(* IEC 61131-3 sources: daoli-st-library/DL_Motion (part 11) *)

(* ---- FB_DL_CamOverrideTrim.st ---- *)
(*
  FB_DL_CamOverrideTrim  —  凸轮运行中动态修调（幅值/相位偏置实时叠加）/ In-run cam dynamic override trim
  分类 Category : DL_Motion
  码位 Code     : 16#04_0_A6
  段位说明      : 04_0 段占至 A5，A6 格空穴，本件启用 A6 格
  版本 Version  : 1.0.1
  来源 Source   : t1-6-plcopen — T1-6 行待挖项「凸轮动态修调」落地
  溯源 Origin   : clean-room 实现，未复制任何源码行
  功能 Function : 1) 不重选表、不脱耦：在 FC_DL_CamTableInterp 表插值输出上实时叠加修调；
                  2) 相位偏置 fPhaseTrim：主轴位置先叠加相位偏置再查表（fMasterEff = fMasterPos + fPhaseTrim），
                  周期模式下按 fPeriod 取模回界，非周期模式下越界按表界钳制（bInRange 反映真实界内性）；
                  3) 幅值偏置 fAmpTrim：从轴输出直接叠加（fSlaveTrimmed = fSlavePos + fAmpTrim）；
                  4) bTrimFreeze 电平冻结修调：冻结拍输出纯表值（修调增量记忆保留，解冻即恢复）。
  边界 Boundary : ① 本件只做输出叠加，不写轴命令、不下使能，凸轮耦合本体由上层承载；
                  ② 与 FC_DL_CamTableInterp（表插值原子）与 FB_DL_ElectronicCam（耦合本体）分工明确；
                  ③ 修调量非有限防御：NaN/Inf 保持上次有效修调值（增量语义不突变）；
                  ④ 无 CASE 主状态机（变换型 FB）：无相位迁移，无跨相 TON 复用问题；
                  ⑤ 本件每拍必须调用一次（无定时器/边沿实例，跳拍仅导致输出陈旧，无隐藏状态损坏）。
  依赖 Depends  : I_DL_MotionAxis（注入，不实例化，只读 fPosition）；
                  FC_DL_CamTableInterp（函数调用，aCam 固定上界透传 + uPointCnt 显式点数）；ST_DL_CamPoint（库内既有结构）
  码表 Error codes（本件格 04_0_A6，子码步进 +0x100）:
    16#0004_01A6 信息级：修调量非有限已保持上次有效值（继续输出，不中断）
    16#0004_02A6 信息级：插值件报错码透传（表非法/越界，本件输出钳界表值）
    16#0004_03A6 信息级：冻结使能中（bTrimFreeze = TRUE，输出纯表值）

  修订历史 Revision :
    2026-11-19  v1.0.0  R39 首版（批次 2 · 序号 7）
    2026-11-23  v1.0.1  R75 适配插值件显式点数字段：aCam 改固定上界 ARRAY[1..200]，
                        增输入 uPointCnt 透传（解 VLA 透传 E037）
*)

FUNCTION_BLOCK FB_DL_CamOverrideTrim
VAR_INPUT
    bEnable     : BOOL := FALSE;      // 使能，FALSE 时输出纯表值（修调旁路）/ Enable, FALSE bypasses trim
    bTrimFreeze : BOOL := FALSE;      // 修调冻结，电平有效：冻结拍输出纯表值 [-] / Trim freeze, level active
    fAmpTrim    : REAL := 0.0;        // 幅值偏置 [mm]，直接叠加从轴输出 / Amplitude trim, added to slave output
    fPhaseTrim  : REAL := 0.0;        // 相位偏置 [mm]，叠加主轴位置后查表 / Phase trim, added to master position
    bPeriodic   : BOOL := FALSE;      // 周期模式使能（与插值件同口径透传）/ Periodic mode, passed to interpolator
    fPeriod     : LREAL := 360.0;     // 周期模式主轴周期 [mm]，域 > 0 / Master period for periodic mode
    bReset      : BOOL := FALSE;      // 修调复位，上升沿清修调保持值（重新从 0 起）/ Trim reset, rising edge clears hold
    uPointCnt   : UINT := 100;        // 凸轮表有效点数，域 [2,200]，透传插值件 [点] / Valid table point count, passthrough to interpolator
END_VAR
VAR_OUTPUT
    fSlaveBase    : LREAL;            // 纯表值输出 [mm]（未叠加修调）/ Pure table output without trim
    fSlaveTrimmed : LREAL;            // 修调后从轴输出 [mm] / Trimmed slave output
    bInRange      : BOOL;             // 有效主轴位置在表界内 [-] / Effective master position within table range
    bTrimActive   : BOOL;             // 修调实际生效中（使能且未冻结且偏置非零）/ Trim actually active
    bClampEdge    : BOOL;             // 相位偏置越表界被钳制（非周期模式）/ Phase trim clamped at table edge
    uErrorId      : UDINT;            // 事件码，0 = 无事件（本件码均信息级瞬时）/ Event code, transient info only
END_VAR
VAR_IN_OUT
    iAxis : I_DL_MotionAxis;          // 主轴引用（注入，不实例化，只读位置）/ Master axis reference, position read-only
    aCam  : ARRAY[1..200] OF ST_DL_CamPoint; // 凸轮表透传（固定上界，下标 1..uPointCnt 有效，须按 fMaster 升序）/ Cam table passed through, fixed bound
END_VAR
VAR
    rtReset      : R_TRIG;            // 修调复位沿实例，主体首部无条件刷新 / Trim reset edge instance
    _bInRangeInt : BOOL;              // 插值件表界内标志内部镜像（段 3 每拍接收，直赋出口）[-] / Interp in-range mirror, received every scan in seg 3
    fAmpTrimEff  : REAL := 0.0;       // 生效幅值偏置 [mm]（非有限保持载体）/ Effective amplitude trim with hold
    fPhaseTrimEff: REAL := 0.0;       // 生效相位偏置 [mm]（非有限保持载体）/ Effective phase trim with hold
    fMasterEff   : LREAL;             // 修调后有效主轴位置 [mm] / Effective master position after phase trim
    fSlavePos    : LREAL;             // 插值件从轴输出 [mm] / Interpolator slave output
    eInterpErr   : UDINT;             // 插值件本拍错误码透传 / Interpolator error code passthrough
    bDefend      : BOOL;              // 本拍非有限防御触发标志 / Non-finite defense triggered this cycle
END_VAR
VAR CONSTANT
    DL_COT_INF_CAP : LREAL := 1.0E15;   // 非有限值筛查幅值上限 / Non-finite screening cap
END_VAR

(* —— 段 0：边沿实例无条件周期刷新（R7 红线） —— *)
rtReset(CLK := bReset);                 // 修调复位沿刷新，每拍必调

(* —— 段 1：修调量非有限防御（NaN/Inf 保持上次有效值；复位沿清保持） —— *)
bDefend := FALSE;                       // 防御标志预清零
IF (fAmpTrim <> fAmpTrim) OR (ABS(fAmpTrim) > DL_COT_INF_CAP) OR ((fAmpTrim - fAmpTrim) <> 0.0) THEN
    bDefend := TRUE;                    // 幅值偏置非有限：保持上次有效
ELSE
    fAmpTrimEff := fAmpTrim;            // 有效值入保持载体
END_IF
IF (fPhaseTrim <> fPhaseTrim) OR (ABS(fPhaseTrim) > DL_COT_INF_CAP) OR ((fPhaseTrim - fPhaseTrim) <> 0.0) THEN
    bDefend := TRUE;                    // 相位偏置非有限：保持上次有效
ELSE
    fPhaseTrimEff := fPhaseTrim;        // 有效值入保持载体
END_IF
IF rtReset.Q THEN
    fAmpTrimEff := 0.0;                 // 复位沿：幅值修调归零
    fPhaseTrimEff := 0.0;               // 复位沿：相位修调归零
END_IF

(* —— 段 2：相位偏置叠加（主轴位置先偏置，周期模式取模回界） —— *)
IF bPeriodic AND (fPeriod > 0.0) THEN
    fMasterEff := iAxis.fPosition + fPhaseTrimEff;              // 叠加相位偏置
    fMasterEff := fMasterEff - TRUNC(fMasterEff / fPeriod) * fPeriod;   // 取模回界（分母已闸 > 0）
    IF fMasterEff < 0.0 THEN
        fMasterEff := fMasterEff + fPeriod;                     // 负模回正（保持 [0, fPeriod) 域）
    END_IF
    bClampEdge := FALSE;                                        // 周期模式无表界钳制概念
ELSE
    fMasterEff := iAxis.fPosition + fPhaseTrimEff;              // 非周期：直接叠加（界内性由插值件判）
    bClampEdge := FALSE;                                        // 钳制判定由插值件 bInRange 承载
END_IF

(* —— 段 3：调表插值原子（每拍一次；错误码透传） —— *)
FC_DL_CamTableInterp(fMasterPos := fMasterEff,      // 有效主轴位置（已含相位偏置）
                     bPeriodic := bPeriodic,        // 周期模式透传
                     fPeriod := fPeriod,            // 周期透传
                     uPointCnt := uPointCnt,        // 显式点数透传（R75 口径）/ Explicit point count passthrough
                     aCam := aCam,                  // 凸轮表透传（固定上界数组引用）
                     fSlavePos => fSlavePos,        // 从轴表值输出
                     bInRange => _bInRangeInt,      // 表界内标志输出（内部镜像）/ In-range flag to internal mirror
                     eErr => eInterpErr);           // 插值件错误码输出
fSlaveBase := fSlavePos;                            // 纯表值镜像
bInRange := _bInRangeInt;                           // 表界内标志出口每拍直赋（语义：有效主轴位置在凸轮表界内为 TRUE）/ In-range outlet assigned every scan

(* —— 段 4：幅值修调叠加与使能门控 —— *)
IF bEnable AND (NOT bTrimFreeze) THEN
    fSlaveTrimmed := fSlaveBase + fAmpTrimEff;      // 修调生效：表值 + 幅值偏置
    bTrimActive := (fAmpTrimEff <> 0.0) OR (fPhaseTrimEff <> 0.0);   // 修调非零即生效中
ELSE
    fSlaveTrimmed := fSlaveBase;                    // 旁路/冻结：输出纯表值（修调保持值不丢）
    bTrimActive := FALSE;
END_IF

(* —— 段 5：事件码合成（信息级瞬时，无锁存） —— *)
uErrorId := 16#0000_0000;               // 缺省无事件
IF bDefend THEN
    uErrorId := 16#0004_01A6;           // 信息级：修调量非有限已保持
ELSIF eInterpErr <> 0 THEN
    uErrorId := 16#0004_02A6;           // 信息级：插值件错误码透传
END_IF
IF bTrimFreeze AND bEnable THEN
    uErrorId := 16#0004_03A6;           // 信息级：冻结使能中（覆盖优先级最低，放最后）
END_IF

END_FUNCTION_BLOCK

(* ---- FB_DL_CamPhaseTrim.st ---- *)
(*
    FB_DL_CamPhaseTrim —— 凸轮相位在线修调
    ------------------------------------------------------------------
    分类      : DL_Motion / Cam
    前缀      : FB_DL_
    版本      : 1.0.0
    溯源      : 只借「凸轮相位可在线修调属运动层能力」的公开语义与运动层组织事实；
                限速率渐进、标记沿一次性受理、相位归一的禁 MOD 写法、错误分级与
                码位 100% 自有；本件不自造轴状态、不内联凸轮算法（组合调用上层凸轮件）；
                clean-room 重写，未复制任何闭源厂商源码
    平台      : 纯 IEC 61131-3，CODESYS V3.5+ / TwinCAT 3 / InoProShop 通用
    作者      : 道莅代码库 · PLC编程专家（R19）
    ------------------------------------------------------------------
    功能说明  : 运行中在线修调凸轮相位，输出一个相位偏移量注入凸轮件的相位输入
                （组合而非内联：可依赖低层，但不复制低层）。现场语义是飞剪/横切/贴标的
                切点对位——用色标或标记传感器测到实际相位偏差后一点点修，修的过程必须
                限速率，突变等于给机械一个冲击。
                核心防御：① 相位限幅越域（> 180°）或速率越域即故障级 02E1 并冻结修调——
                   相位限幅 0 会让修调永久卡住、太大等于允许突变；
                ② 一次性标记补偿每标记沿只受理一次，且必须在 bMarkArmed（上一拍已复位）
                   时才受理——否则高频标记会在一拍内累加成大跳变（本件最高危点）；
                ③ 相位归一用条件加减，禁浮点 MOD；
                ④ 指令或补偿量非有限即故障级并保持末次偏移——归 0 会让切点瞬间错位切出废品；
                ⑤ bReset 立即清偏移（唯一允许跳变的路径，检修专用）。
                职责边界：凸轮曲线求值归电子凸轮件，本件只出相位偏移量。
    错误码    : 16#0004_01CF 目标偏移超限已钳位 / 单次标记补偿已生效——信息级，正常防御
                16#0004_01D0 预留禁用（信息级，不得挪用）
                16#0004_02E1 限幅、速率或采样周期参数非法——故障级，修调冻结且偏移保持
                16#0004_02E2 指令或补偿量非有限——故障级，偏移保持末次有效
                16#0004_02E3 状态机落 ELSE 兜底（非法状态）——故障级，回 eIdle 并保持偏移
    码位总账  : 16#0004_01CF 用 / 16#0004_01D0 预留 ｜ 16#0004_02E1 用 / 16#0004_02E2 用 / 16#0004_02E3 用
    状态机    : E_DL_TrimState（eIdle / eRamping / eHold / eFault）四态，CASE 含 ELSE 兜底，
                ELSE 回 eIdle 并置故障级 02E3；失能时目标归 0 并按限速率回零。
    采样约定  : fbTrigReset / fbTrigMark 在本体首部无条件刷新，绝不放入 IF 或 CASE；
                速率步长由 tSampleTime 引脚换算，首拍步长按引脚值直接给出（无历史依赖）。
    修订记录  : 2026-11-16 v1.0.0 首次入库（R19）
*)

(*
    枚举 : E_DL_TrimState —— 相位修调状态（本文件为全库唯一属主）
*)
TYPE E_DL_TrimState :
(
    eIdle    := 0,                            // 空闲：偏移按限速率回零 / idle, the offset ramps back to zero
    eRamping := 1,                            // 趋近：向目标偏移逼近 / ramping towards the target offset
    eHold    := 2,                            // 保持：已到目标，仅受标记补偿影响 / holding at the target
    eFault   := 3                             // 故障：修调冻结，偏移保持 / fault, the trim is frozen and the offset held
);
END_TYPE

FUNCTION_BLOCK FB_DL_CamPhaseTrim
VAR_INPUT
    bEnable         : BOOL;                   // 使能，FALSE 偏移按限速率归 0 / enable, FALSE ramps the offset back to zero
    bReset          : BOOL;                   // 复位，上升沿立即清偏移（检修专用，会跳变）/ reset, rising edge clears the offset at once, maintenance only
    fPhaseOffsetCmd : REAL := 0.0;            // 目标相位偏移 [deg]，范围 -180.0~180.0 / target phase offset [deg], range -180.0~180.0
    fRateMax        : REAL := 30.0;           // 偏移变化率上限 [deg/s]，范围 0.1~3600.0 / maximum offset rate [deg/s], range 0.1~3600.0
    fPhaseLimit     : REAL := 90.0;           // 偏移绝对值上限 [deg]，范围 1.0~180.0 / absolute offset limit [deg], range 1.0~180.0
    bTrimOnMark     : BOOL := FALSE;          // TRUE = 叠加标记沿的一次性补偿 / TRUE adds the one-shot mark correction
    fMarkCorrection : REAL := 0.0;            // 单次标记补偿量 [deg]，范围 -10.0~10.0 / one-shot mark correction [deg], range -10.0~10.0
    bMarkPulse      : BOOL := FALSE;          // 标记传感器脉冲（上升沿有效）/ mark sensor pulse, rising edge valid
    tSampleTime     : TIME := T#10MS;         // 采样周期 [ms]，范围 1~1000 / sample time [ms], range 1~1000
END_VAR
VAR_OUTPUT
    fPhaseOffset    : REAL;                   // 实际输出相位偏移（注入凸轮件）[deg] / actual phase offset injected into the cam block [deg]
    bTrimming       : BOOL;                   // 正在趋近目标 / ramping towards the target
    bLimited        : BOOL;                   // 受速率或幅值限制 / limited by the rate or the magnitude
    uMarkCount      : UDINT;                  // 已受理的标记补偿次数，饱和 [次] / accepted mark corrections, saturating [times]
    eErr            : UDINT;                  // 错误码，0=正常 / error id, 0=ok
    bError          : BOOL;                   // 故障标志，eErr 为故障级时 TRUE / error flag, TRUE on fault-level eErr
END_VAR
VAR
    fbTrigReset     : R_TRIG;                 // 复位上升沿实例，本体首部无条件刷新 / reset edge instance, refreshed unconditionally
    fbTrigMark      : R_TRIG;                 // 标记上升沿实例，本体首部无条件刷新 / mark edge instance, refreshed unconditionally
    eState          : E_DL_TrimState := eIdle; // 状态机当前态 / current state machine state
    fOffset         : REAL;                   // 内部偏移量 [deg] / internal offset [deg]
    fTarget         : REAL;                   // 限幅后的目标偏移 [deg] / clamped target offset [deg]
    fStep           : REAL;                   // 本拍允许的最大变化量 [deg] / maximum allowed change in this cycle [deg]
    fDtSec          : REAL;                   // 采样周期秒值 [s] / sample time in seconds [s]
    fLimitEff       : REAL;                   // 钳位后的相位限幅 [deg] / clamped phase limit [deg]
    fCorrEff        : REAL;                   // 钳位后的单次补偿量 [deg] / clamped one-shot correction [deg]
    bMarkArmed      : BOOL := TRUE;           // 标记受理武装位（上一拍已复位才受理）/ mark acceptance arming bit, armed only after the pulse is released
    bNonFin         : BOOL;                   // 输入非有限判定标志 / non-finite input flag
    bInit           : BOOL := FALSE;          // 首扫标志，初值 FALSE，判据 NOT bInit / first-scan flag, initial FALSE, tested with NOT
    nDtMs           : DINT;                   // 采样周期毫秒整数 [ms] / sample time in integer milliseconds [ms]
END_VAR
VAR CONSTANT
    DL_CPT_LIMIT_MAX : REAL := 180.0;         // 相位限幅上限（半周）[deg] / phase limit upper bound, half a revolution [deg]
    DL_CPT_LIMIT_MIN : REAL := 1.0;           // 相位限幅下限 [deg] / phase limit lower bound [deg]
    DL_CPT_RATE_MAX  : REAL := 3600.0;        // 速率上限 [deg/s] / rate upper bound [deg/s]
    DL_CPT_RATE_MIN  : REAL := 0.1;           // 速率下限 [deg/s] / rate lower bound [deg/s]
    DL_CPT_MARK_MAX  : REAL := 10.0;          // 单次补偿量绝对值上限 [deg] / absolute one-shot correction bound [deg]
    DL_CPT_DT_MAX    : TIME := T#1S;          // 采样周期上限 [ms] / sample time upper bound [ms]
    DL_CPT_DT_MIN    : TIME := T#1MS;         // 采样周期下限 [ms] / sample time lower bound [ms]
    DL_FLOAT_EPS     : REAL := 1.0E-6;        // 浮点判等容差 [无量纲] / float equality tolerance [dimensionless]
    DL_CPT_FULL_TURN : REAL := 360.0;         // 一整周 [deg] / one full revolution [deg]
    DL_CPT_HALF_TURN : REAL := 180.0;         // 半周 [deg] / half a revolution [deg]
    DL_CPT_MS_PER_S  : REAL := 1000.0;        // 毫秒到秒换算因子 [ms/s] / milliseconds per second [ms/s]
    DL_CPT_INF_GUARD : REAL := 1.0E38;        // 非有限幅值判定阈值 [无量纲] / non-finite magnitude guard [dimensionless]
    DL_CPT_CNT_MAX   : UDINT := 16#FFFF_FFFE; // 标记次数饱和值 [次] / mark counter saturation value [times]
    DL_CPT_ZERO      : REAL := 0.0;           // 零值常量，避免裸字面量 [deg] / zero constant, avoids a bare literal [deg]
END_VAR

// 段 1｜边沿实例无条件周期刷新（红线：严禁放入条件分支）/ segment 1, unconditional edge refresh
fbTrigReset(CLK := bReset);
fbTrigMark(CLK := bMarkPulse);

// 段 2｜输出与错误状态预置 / segment 2, preset outputs and status
eErr := 0;                                    // 预置无错误 / preset no error
bError := FALSE;                              // 预置无故障 / preset no fault
bTrimming := FALSE;                           // 预置未趋近 / preset not ramping
bLimited := FALSE;                            // 预置未受限 / preset not limited

// 段 3｜首扫初始化（唯一合法范式：初值 FALSE，判据 NOT bInit）/ segment 3, first-scan initialisation
IF NOT bInit THEN
    fOffset := DL_CPT_ZERO;                   // 首扫偏移归 0，避免未定值上电冲击 / the offset starts at zero, no undefined jump at power up
    uMarkCount := 0;                          // 标记计数清零 / clear the mark counter
    bInit := TRUE;                            // 首扫只做一次 / first scan runs once only
END_IF

// 段 4｜参数闸（限幅、速率、采样周期，任一非法即冻结修调）/ segment 4, parameter gate freezes the trim
IF (fPhaseLimit < DL_CPT_LIMIT_MIN) OR (fPhaseLimit > DL_CPT_LIMIT_MAX)
   OR (fRateMax < DL_CPT_RATE_MIN) OR (fRateMax > DL_CPT_RATE_MAX)
   OR (tSampleTime < DL_CPT_DT_MIN) OR (tSampleTime > DL_CPT_DT_MAX) THEN
    eErr := 16#0004_02E1;                     // 参数非法故障码 / illegal parameter fault id
    bError := TRUE;                           // 置故障标志 / raise the error flag
    eState := eFault;                         // 落故障态，修调冻结 / enter the fault state, the trim is frozen
    fPhaseOffset := fOffset;                  // 偏移保持，绝不归 0 / hold the offset, never reset it to zero
    RETURN;                                   // 故障级提前返回 / early return on fault
END_IF

// 段 5｜输入非有限闸：偏移保持末次有效（归 0 会瞬间错位切出废品）/ segment 5, non-finite gate holds the offset
bNonFin := (fPhaseOffsetCmd <> fPhaseOffsetCmd) OR (fMarkCorrection <> fMarkCorrection)
        OR (fPhaseOffsetCmd > DL_CPT_INF_GUARD) OR (fPhaseOffsetCmd < -DL_CPT_INF_GUARD); // 非有限判定 / non-finite detection
IF bNonFin THEN
    eErr := 16#0004_02E2;                     // 指令非有限故障码 / non-finite command fault id
    bError := TRUE;                           // 置故障标志 / raise the error flag
    eState := eFault;                         // 落故障态 / enter the fault state
    fPhaseOffset := fOffset;                  // 保持末次有效偏移 / hold the last valid offset
    RETURN;                                   // 故障级提前返回 / early return on fault
END_IF

// 段 5｜域钳位（限幅、补偿量各自收敛，钳位本身不置码）/ segment 5, domain clamp
fLimitEff := MIN(MAX(fPhaseLimit, DL_CPT_LIMIT_MIN), DL_CPT_LIMIT_MAX);   // 相位限幅收敛 [deg] / converge the phase limit [deg]
fCorrEff := MIN(MAX(fMarkCorrection, -DL_CPT_MARK_MAX), DL_CPT_MARK_MAX); // 单次补偿收敛到 ±10 deg / converge the one-shot correction
nDtMs := TIME_TO_DINT(tSampleTime);           // 采样周期整数毫秒 [ms] / sample time in integer milliseconds [ms]
fDtSec := DINT_TO_REAL(nDtMs) / DL_CPT_MS_PER_S; // 换算为秒，除子为常量 [s] / convert to seconds, the divisor is a constant [s]
fStep := fRateMax * fDtSec;                   // 本拍允许的最大变化量 [deg] / maximum allowed change in this cycle [deg]

// 段 6｜目标偏移 = 指令限幅 / segment 6, target offset from the clamped command
fTarget := MIN(MAX(fPhaseOffsetCmd, -fLimitEff), fLimitEff); // 目标双侧钳位 [deg] / clamp the target on both sides [deg]
IF ABS(fPhaseOffsetCmd) > fLimitEff THEN
    eErr := 16#0004_01CF;                     // 信息级：目标偏移超限已钳位 / info level, the target was clamped
END_IF

// 段 7｜标记沿一次性补偿（最高危点：每沿只受理一次，且需武装位）/ segment 7, one-shot mark correction
IF NOT bMarkPulse THEN
    bMarkArmed := TRUE;                       // 脉冲释放即重新武装 / re-arm once the pulse is released
END_IF
IF fbTrigMark.Q AND bTrimOnMark AND bMarkArmed THEN
    bMarkArmed := FALSE;                      // 受理后立即解除武装，防同拍累加 / disarm immediately so no accumulation can happen in one cycle
    fTarget := MIN(MAX(fTarget + fCorrEff, -fLimitEff), fLimitEff); // 叠加补偿并限幅 [deg] / add the correction and clamp [deg]
    IF uMarkCount < DL_CPT_CNT_MAX THEN
        uMarkCount := uMarkCount + 1;         // 饱和计数 / saturating count
    END_IF
    eErr := 16#0004_01CF;                     // 信息级：单次标记补偿已生效 / info level, the one-shot correction was applied
END_IF

// 段 8｜复位沿：立即清偏移（唯一允许跳变的路径，检修专用）/ segment 8, reset clears the offset at once
IF fbTrigReset.Q THEN
    fOffset := DL_CPT_ZERO;                   // 检修专用清偏移 / maintenance only, clear the offset
    bLimited := FALSE;                        // 清限幅标志 / clear the limited flag
END_IF

// 段 9｜失能：目标归 0，按限速率回零 / segment 9, disabling ramps the target back to zero
IF NOT bEnable THEN
    fTarget := DL_CPT_ZERO;                   // 目标归 0 / the target returns to zero
END_IF

// 段 10｜状态机（含 ELSE 兜底）/ segment 10, state machine with ELSE fallback
CASE eState OF
    eIdle:
        IF ABS(fTarget - fOffset) > fStep THEN
            eState := eRamping;               // 偏离超过一步即进入趋近态 / a deviation beyond one step enters the ramping state
        ELSE
            eState := eHold;                  // 否则直接保持 / otherwise hold at once
        END_IF

    eRamping:
        IF ABS(fTarget - fOffset) <= fStep THEN
            eState := eHold;                  // 进入一步之内即趋近完成 / inside one step the ramp is finished
        END_IF

    eHold:
        IF ABS(fTarget - fOffset) > fStep THEN
            eState := eRamping;               // 新指令或标记补偿把偏差拉大即重新趋近 / a new command or correction restarts the ramp
        END_IF

    eFault:
        fPhaseOffset := fOffset;              // 故障态偏移保持 / hold the offset in the fault state

ELSE
    eErr := 16#0004_02E3;                     // 故障级：非法状态兜底 / fault level, illegal state fallback
    bError := TRUE;                           // 置故障标志 / raise the error flag
    eState := eIdle;                          // 回空闲态 / fall back to idle
    fPhaseOffset := fOffset;                  // 保持偏移，绝不清零 / hold the offset, never clear it
END_CASE

// 段 11｜限速率推进（每拍最多变化 fStep，禁浮点 MOD 的相位归一）/ segment 11, rate limited advance
IF eState <> eFault THEN
    IF fOffset > (fTarget + fStep) THEN
        fOffset := fOffset - fStep;           // 正向逼近 / approach from above
        bLimited := TRUE;                     // 标记速率受限 / flag the rate limit
        bTrimming := TRUE;                    // 正在趋近 / ramping
    ELSIF fOffset < (fTarget - fStep) THEN
        fOffset := fOffset + fStep;           // 负向逼近 / approach from below
        bLimited := TRUE;                     // 标记速率受限 / flag the rate limit
        bTrimming := TRUE;                    // 正在趋近 / ramping
    ELSE
        fOffset := fTarget;                   // 进入一步之内即直接到位 / snap into place once inside one step
        bTrimming := FALSE;                   // 到位即不再趋近 / no longer ramping
    END_IF

    // 段 12｜幅值限幅（双侧，超限置受限标志）/ segment 12, two-sided magnitude clamp
    IF fOffset > fLimitEff THEN
        fOffset := fLimitEff;                 // 正向限幅 / clamp the positive side
        bLimited := TRUE;                     // 标记幅值受限 / flag the magnitude limit
    ELSIF fOffset < -fLimitEff THEN
        fOffset := -fLimitEff;                // 负向限幅 / clamp the negative side
        bLimited := TRUE;                     // 标记幅值受限 / flag the magnitude limit
    END_IF

    // 段 13｜相位归一（条件加减，禁浮点 MOD）/ segment 13, phase normalisation without a floating point MOD
    IF fOffset > DL_CPT_HALF_TURN THEN
        fOffset := fOffset - DL_CPT_FULL_TURN; // 超半周折回一周 / fold back one revolution
    ELSIF fOffset < -DL_CPT_HALF_TURN THEN
        fOffset := fOffset + DL_CPT_FULL_TURN; // 低于负半周折回一周 / fold forward one revolution
    END_IF
END_IF

// 段 14｜发布结果 / segment 14, publish the result
fPhaseOffset := fOffset;                      // 输出实际偏移（回零过程亦发布真实值）[deg] / publish the actual offset, including the ramp back to zero [deg]
END_FUNCTION_BLOCK

(* ---- FB_DL_CamSlavePhaseOffsetSeq.st ---- *)
(*
  Name: FB_DL_CamSlavePhaseOffsetSeq
  Category: DL_Motion
  Version: 1.0.0
  Round: R89 / 2026-11-25
  开源溯源：clean-room 自研（族 运动同步控制，ST 开源生态实测 0 命中，无外部代码引入）
  功能：凸轮从动相位偏置在线切换：偏置斜坡 + 接合点判定，非接合点/关键区一律拒绝并给出 ENUM 原因。
  边界条件：① 五浮点入参全部过非有限闸，配置越域即锁故障（eFault），拒因出口同拍置 eCfgBad；
            ② 切换许可四项与门：使能、啮合（xInMesh）、非关键区、目标在 ±90° 内；任一不满足即拒并锁拒因；
            ③ 关键区（接合禁区）定义为相位 0~20° 与 340~360° 两段（相位按 0~360 口径输入）；
            ④ 斜坡起点取实测偏置 fOffsetActDeg，避免切换瞬间偏置跳变；步长 = fRampDegPerS × fCycleS；
            ⑤ 斜坡中若啮合丢失立即中止（拒因 eNotInMesh），已走偏置保持，不再回退；
            ⑥ 故障解除唯一路径：故障相内 xEnable 释放（R152），清锁存回 eIdle。
  状态机：eIdle / eHold / eRamp / eFault（CASE 含 ELSE 兜底）。
  量纲自证：°/s × s = °；偏置与目标同为 °，容差比较同量纲。
*)
TYPE E_DL_CspoPhase :
(
    eIdle  := 0,        (* 待机：未使能 / Idle, not enabled *)
    eHold  := 10,       (* 保持相：偏置保持，等切换申请 / Hold, waiting switch request *)
    eRamp  := 20,       (* 斜坡相：偏置向目标推进 / Ramping offset to target *)
    eFault := 90        (* 故障相：配置越域锁存 / Fault, configuration latched *)
);
END_TYPE
TYPE E_DL_CspoReject :
(
    eNone       := 0,   (* 无拒绝（最近一次切换被接受） / No rejection, last switch accepted *)
    eNotEnabled := 1,   (* 拒绝：未使能 / Rejected, not enabled *)
    eNotInMesh  := 2,   (* 拒绝：凸轮未啮合（或斜坡中脱啮） / Rejected, cam not in mesh *)
    eKeyZone    := 3,   (* 拒绝：处于关键区（接合禁区） / Rejected, inside key zone *)
    eTargetLim  := 4,   (* 拒绝：目标偏置超 ±90° / Rejected, target beyond limit *)
    eCfgBad     := 5    (* 拒绝：组态非法（非有限或越域） / Rejected, bad configuration *)
);
END_TYPE

FUNCTION_BLOCK FB_DL_CamSlavePhaseOffsetSeq
VAR_INPUT
    xEnable : BOOL;             (* 使能 [-] Enable *)
    xSwitchCmd : BOOL;          (* 切换申请（上升沿有效） [-] Switch request, rising edge *)
    fPhaseActDeg : REAL;        (* 凸轮实际相位（0~360） [°] Cam actual phase [deg] *)
    fOffsetTargetDeg : REAL;    (* 目标偏置 [°] Target offset [deg] *)
    fOffsetActDeg : REAL;       (* 实测偏置（斜坡起点） [°] Actual offset [deg] *)
    fRampDegPerS : REAL;        (* 偏置斜坡速率 [°/s] Offset ramp rate [deg/s] *)
    xInMesh : BOOL;             (* 凸轮啮合反馈 [-] Cam in mesh *)
    fCycleS : REAL;             (* 扫描周期 [s] Scan cycle [s] *)
END_VAR
VAR_OUTPUT
    fOffsetOutDeg : REAL;       (* 偏置输出（斜坡后） [°] Offset output [deg] *)
    eState : E_DL_CspoPhase;    (* 当前相 [-] Present phase *)
    xApplyDone : BOOL;          (* 切换完成单拍脉冲 [-] One-scan apply done *)
    xRejectReason : E_DL_CspoReject;    (* 最近一次切换的拒绝原因 [-] Reject reason *)
    xFault : BOOL;              (* 故障锁存标志 [-] Fault latched *)
END_VAR
VAR
    _eState : E_DL_CspoPhase := E_DL_CspoPhase.eIdle;  (* 内部相（CASE 唯一写入目标） [-] Internal phase *)
    _eReject : E_DL_CspoReject := E_DL_CspoReject.eNone;   (* 拒因锁存 [-] Reject reason latch *)
    _bInit : BOOL := FALSE;         (* 首扫初始化标志 [-] First-scan init flag *)
    _bFaultLatch : BOOL := FALSE;   (* 故障锁存位 [-] Fault latch *)
    _bApply : BOOL := FALSE;        (* 单拍完成标志（段 2 预清） [-] One-scan apply flag *)
    _bRampReq : BOOL := FALSE;      (* 当拍切换受理标志（段 2 预清） [-] Switch accepted flag *)
    _bCfgBad : BOOL := FALSE;       (* 配置非法当拍量 [-] Configuration bad *)
    _bKeyZone : BOOL := FALSE;      (* 关键区判据 [-] Inside key zone *)
    _fOut : REAL := 0.0;            (* 偏置输出保持量 [°] Offset output hold [deg] *)
    _fStep : REAL := 0.0;           (* 单拍斜坡步长 [°] Ramp step [deg] *)
    _fCy : REAL := 0.01;            (* 当拍有效周期 [s] Effective cycle [s] *)
    rtSwitch : R_TRIG;              (* 切换沿（段 1 无条件调用） / Switch edge *)
END_VAR
VAR CONSTANT
    DL_CSPO_TOL : REAL := 0.05;     (* 偏置到位容差 [°] Offset tolerance [deg] *)
    DL_CSPO_MAX : REAL := 90.0;     (* 目标偏置工程限 [°] Target offset limit [deg] *)
    DL_CSPO_KEY_HALF : REAL := 20.0;(* 关键区半宽（0~20 与 340~360） [°] Key zone half width [deg] *)
    DL_CSPO_FULL : REAL := 360.0;   (* 整转角度 [°] Full revolution [deg] *)
    DL_CSPO_CYDEF : REAL := 0.01;   (* 缺省扫描周期 [s] Default scan cycle [s] *)
    DL_CSPO_RATE_MIN : REAL := 1.0; (* 斜坡速率下限 [°/s] Ramp rate floor [deg/s] *)
    DL_CSPO_RATE_MAX : REAL := 720.0;   (* 斜坡速率上限 [°/s] Ramp rate ceiling [deg/s] *)
END_VAR
(* —— 段 0：非有限闸（NaN 自反 + Inf 差值自减）+ 组态域闸，五浮点入参全枚举（R272） —— *)
_bCfgBad := (fPhaseActDeg <> fPhaseActDeg) OR ((fPhaseActDeg - fPhaseActDeg) <> 0.0)
         OR (fOffsetTargetDeg <> fOffsetTargetDeg) OR ((fOffsetTargetDeg - fOffsetTargetDeg) <> 0.0)
         OR (fOffsetActDeg <> fOffsetActDeg) OR ((fOffsetActDeg - fOffsetActDeg) <> 0.0)
         OR (fRampDegPerS <> fRampDegPerS) OR ((fRampDegPerS - fRampDegPerS) <> 0.0)
         OR (fCycleS <> fCycleS) OR ((fCycleS - fCycleS) <> 0.0)
         OR (fPhaseActDeg < 0.0) OR (fPhaseActDeg > DL_CSPO_FULL)
         OR (fOffsetTargetDeg > DL_CSPO_MAX) OR (fOffsetTargetDeg < (0.0 - DL_CSPO_MAX))
         OR (fOffsetActDeg > DL_CSPO_MAX) OR (fOffsetActDeg < (0.0 - DL_CSPO_MAX))
         OR (fRampDegPerS < DL_CSPO_RATE_MIN) OR (fRampDegPerS > DL_CSPO_RATE_MAX);
(* 关键区判据：相位 0~20° 或 340~360° 为接合禁区 *)
_bKeyZone := (fPhaseActDeg <= DL_CSPO_KEY_HALF)
          OR (fPhaseActDeg >= (DL_CSPO_FULL - DL_CSPO_KEY_HALF));
(* 周期派生：非法周期取 10 ms 缺省 *)
IF (fCycleS > 0.0) AND (fCycleS <= 1.0) THEN
    _fCy := fCycleS;
ELSE
    _fCy := DL_CSPO_CYDEF;
END_IF
(* 首扫初始化：偏置输出以实测偏置播种，避免首拍跳变（R310） *)
IF NOT _bInit THEN
    (* 播种前非有限闸：NOT(x<=360) 对 NaN 为真，防 NaN 播种后永久冻结 *)
    IF (fOffsetActDeg <= 360.0) AND (fOffsetActDeg >= -360.0) THEN
        _fOut := fOffsetActDeg;
    ELSE
        _fOut := 0.0;                       (* 实测偏置无效即零播种 / Seed zero on invalid actual *)
    END_IF
    _bInit := TRUE;
END_IF
(* —— 段 1：切换沿无条件刷新（R7） —— *)
rtSwitch(CLK := xSwitchCmd);
(* —— 段 2：单拍量预清 —— *)
_bApply := FALSE;
_bRampReq := FALSE;
(* —— 段 3：切换受理校验（拒因唯一出口，逐项归因互不共用成员，R190） —— *)
IF rtSwitch.Q THEN
    IF _bCfgBad THEN
        _eReject := E_DL_CspoReject.eCfgBad;        (* 组态非法 / Bad configuration *)
    ELSIF NOT xEnable THEN
        _eReject := E_DL_CspoReject.eNotEnabled;    (* 未使能 / Not enabled *)
    ELSIF NOT xInMesh THEN
        _eReject := E_DL_CspoReject.eNotInMesh;     (* 未啮合 / Not in mesh *)
    ELSIF _bKeyZone THEN
        _eReject := E_DL_CspoReject.eKeyZone;       (* 关键区 / Key zone *)
    ELSIF (fOffsetTargetDeg > DL_CSPO_MAX) OR (fOffsetTargetDeg < (0.0 - DL_CSPO_MAX)) THEN
        _eReject := E_DL_CspoReject.eTargetLim;     (* 目标越限 / Target over limit *)
    ELSE
        _eReject := E_DL_CspoReject.eNone;          (* 受理 / Accepted *)
        _bRampReq := TRUE;
    END_IF
END_IF
(* —— 段 4：故障锁存解除（唯一路径 = 故障相内 xEnable 释放，R152） —— *)
IF _bFaultLatch AND (NOT xEnable) THEN
    _bFaultLatch := FALSE;                      (* 清锁存 / Clear latch *)
    _eState := E_DL_CspoPhase.eIdle;            (* 迁回待机 / Back to idle *)
END_IF
(* —— 段 5：主状态机（ENUM + CASE，ELSE 兜底） —— *)
CASE _eState OF
E_DL_CspoPhase.eIdle:
    IF xEnable AND (NOT _bFaultLatch) THEN
        _fOut := fOffsetActDeg;                 (* 上电取实测偏置为起点 / Seed from actual *)
        _eState := E_DL_CspoPhase.eHold;
    END_IF
E_DL_CspoPhase.eHold:
    _fOut := fOffsetActDeg;                     (* 保持相：偏置跟随实测（外部闭环保持） / Hold *)
    IF NOT xEnable THEN
        _eState := E_DL_CspoPhase.eIdle;
    ELSIF _bRampReq THEN
        _fOut := fOffsetActDeg;                 (* 斜坡起点重置为实测值 / Reset start point *)
        _eState := E_DL_CspoPhase.eRamp;
    END_IF
E_DL_CspoPhase.eRamp:
    _fStep := fRampDegPerS * _fCy;              (* °/s × s = ° / Ramp step *)
    IF NOT xInMesh THEN
        _eReject := E_DL_CspoReject.eNotInMesh; (* 斜坡中脱啮：中止 / Mesh lost, abort *)
        _eState := E_DL_CspoPhase.eHold;
    ELSIF NOT xEnable THEN
        _eState := E_DL_CspoPhase.eIdle;        (* 使能撤销 / Enable dropped *)
    ELSIF _fOut < (fOffsetTargetDeg - DL_CSPO_TOL) THEN
        _fOut := _fOut + _fStep;
        IF _fOut > fOffsetTargetDeg THEN
            _fOut := fOffsetTargetDeg;          (* 上钳 / Upper clamp *)
        END_IF
    ELSIF _fOut > (fOffsetTargetDeg + DL_CSPO_TOL) THEN
        _fOut := _fOut - _fStep;
        IF _fOut < fOffsetTargetDeg THEN
            _fOut := fOffsetTargetDeg;          (* 下钳 / Lower clamp *)
        END_IF
    ELSE
        _fOut := fOffsetTargetDeg;              (* 到位落定 / Settle to target *)
        _bApply := TRUE;                        (* 单拍完成（段 2 预清） / One-scan done *)
        _eReject := E_DL_CspoReject.eNone;      (* 本次切换成功，清拒因 / Clear reject *)
        _eState := E_DL_CspoPhase.eHold;
    END_IF
E_DL_CspoPhase.eFault:
    _bKeyZone := (fPhaseActDeg <= DL_CSPO_KEY_HALF)
              OR (fPhaseActDeg >= (DL_CSPO_FULL - DL_CSPO_KEY_HALF));   (* 故障相驻留：判据照算 *)
ELSE
    _bCfgBad := TRUE;                           (* 非法相兜底 / Illegal phase fallback *)
    _eState := E_DL_CspoPhase.eFault;
END_CASE
(* —— 段 6：组态故障统一落地（唯一锁存点 + 同步迁相，R187/R252） —— *)
IF _bCfgBad AND (NOT _bFaultLatch) THEN
    _bFaultLatch := TRUE;                       (* 锁存 / Latch *)
    _eReject := E_DL_CspoReject.eCfgBad;        (* 拒因同拍置 eCfgBad / Reject cause *)
    _eState := E_DL_CspoPhase.eFault;           (* 同步迁相 / Migrate to fault *)
END_IF
(* —— 段 7：统一出口（各出口单点赋值） —— *)
(* 出口非有限闸：偏置输出绝不外泄 NaN / INF *)
IF NOT ((_fOut <= 360.0) AND (_fOut >= -360.0)) THEN
    _fOut := 0.0;                           (* 归零偏置 / Zero offset *)
END_IF
fOffsetOutDeg := _fOut;
eState := _eState;
xApplyDone := _bApply;
xRejectReason := _eReject;
xFault := _bFaultLatch;
END_FUNCTION_BLOCK

(* ---- FB_DL_CamTableLiveTrim.st ---- *)
(*
  Name        : FB_DL_CamTableLiveTrim
  Category    : DL_Motion
  Version     : 1.0.0
  Purpose     : 凸轮表运行中动态修调：指定相位点修调请求经斜坡平滑注入运行表，每次写表随改随验单调性，破坏即回滚本点锁故障；/ Live cam table trim: point trim request ramped smoothly into the running table, monotonicity verified on every write with instant rollback of the point on violation
  溯源        : 借 plcopen-motion 的凸轮动态修调待挖组织，clean-room 实现
  Boundary    : ① 修调注入只允许运行相且主轴相位在目标点 ± 容差窗内（相位闸，容差域 > 0）；
                ② 修调后表值单调性随改随验，破坏单调立即回滚本点至基线快照并锁存故障至复位沿；
                ③ 修调量饱和上限（绝对值钳位）防累计漂移，饱和上限域 > 0；
                ④ 斜坡平滑步长 = 斜坡率 × 周期秒值；非有限修调请求/主轴位置该拍不注入（保持上拍）；
                ⑤ 表经输入输出引用参数注入，内部零表副本（仅存单点基线快照，防两份表失同步）；
                ⑥ 表点数域 2..16，修调点序号越域直接拒绝申请（不置故障，属申请级）。
*)
TYPE E_DL_CltState :
(
    eIdle  := 0,                             (* 未使能 / Disabled *)
    eRun   := 10,                            (* 修调待触发/斜坡注入运行 / Trim running *)
    eFault := 90                             (* 故障锁存相 / Fault latched *)
);
END_TYPE

TYPE E_DL_CltCause :
(
    eNone     := 0,                          (* 无故障成因 / No cause *)
    eCfgIllegal:= 1,                        (* 组态非法：点数/容差/斜率/饱和域越界 / Illegal config *)
    eMonotonic:= 2,                         (* 单调性破坏（回滚 + 锁存，边界②） / Monotonicity violated *)
    ePhaseBad := 3                          (* 非法相位兜底 / Illegal phase fallback *)
);
END_TYPE

FUNCTION_BLOCK FB_DL_CamTableLiveTrim
VAR_INPUT
    fMasterPos: REAL := 0.0;                (* 主轴相位当前位置 [度] / Master phase position *)
    fMasterSpan: REAL := 360.0;             (* 主轴相位量程，域 > 0 [度] / Master span *)
    nPts     : INT := 16;                   (* 表点数，域 2..16 [点] / Table point count *)
    nIdx     : INT := 1;                    (* 修调目标点序号（1 基）[点] / Trim target point index *)
    fTrim    : REAL := 0.0;                 (* 修调请求量（正 = 增大表值）[表值单位] / Trim request amount *)
    fTrimMax : REAL := 1.0;                 (* 单点修调饱和上限，域 > 0 [表值单位] / Trim saturation cap *)
    fRampRate: REAL := 10.0;                (* 斜坡注入率，域 > 0 [表值单位/s] / Ramp rate *)
    fTol     : REAL := 1.0;                 (* 相位闸容差，域 > 0 [度] / Phase gate tolerance *)
    tScan    : TIME := T#10MS;              (* 扫描周期，域 > T#0S [ms] / Scan period *)
    bApply   : BOOL := FALSE;               (* 修调申请，上升沿受理 [-] / Apply request *)
    bEnable  : BOOL := TRUE;                (* 使能 [-] / Enable *)
    bReset   : BOOL := FALSE;               (* 复位命令，上升沿清故障 [-] / Reset command *)
END_VAR
VAR_IN_OUT
    aTable   : ARRAY[1..16] OF REAL;        (* 凸轮表（从动值，零内部副本，边界⑤） / Cam table by reference *)
END_VAR
VAR_OUTPUT
    fApplied : REAL;                        (* 当前已注入修调量（镜像）[表值单位] / Applied trim mirror *)
    bTrimDone: BOOL;                        (* 本拍修调注入完成（单拍脉冲）[-] / Trim done pulse *)
    eState   : E_DL_CltState;               (* 状态出口 / State outlet *)
    eCause   : E_DL_CltCause;               (* 故障成因出口（R190 归因唯一） / Fault cause outlet *)
    bError   : BOOL;                        (* 故障锁存标志 [-] / Fault latch flag *)
END_VAR
VAR
    _eState : E_DL_CltState := E_DL_CltState.eIdle;  (* 内部相位（CASE 唯一写入目标） / Internal phase *)
    _eCause : E_DL_CltCause := E_DL_CltCause.eNone;  (* 故障成因锁存量 / Latched cause *)
    rtApply : R_TRIG;                       (* 申请沿实例，段 0 无条件调用 / Apply edge instance *)
    rtReset : R_TRIG;                       (* 复位沿实例，段 0 无条件调用 / Reset edge instance *)
    _bFault : BOOL;                         (* 故障锁存位 / Latched fault bit *)
    _bCfgBad: BOOL;                         (* 组态非法当拍量 / Illegal config this scan *)
    _bFin   : BOOL;                         (* 主轴相位/修调量有限性当拍量（边界④） / Inputs finiteness *)
    _bDoneI : BOOL;                         (* 完成脉冲内部量（统一出口映射，R187） / Done pulse internal *)
    _bInj   : BOOL;                         (* 斜坡注入进行中标志 / Ramping flag *)
    _nIdxE  : INT;                          (* 受理后生效点序号 [点] / Effective index *)
    _fTarget: REAL;                         (* 饱和钳位后修调目标量 [表值单位] / Clamped trim target *)
    _fApplI : REAL;                         (* 已注入量内部量 [表值单位] / Applied internal *)
    _fBase  : REAL;                         (* 注入起始拍该点基线快照 [表值单位] / Point baseline snapshot *)
    _fStep  : REAL;                         (* 本拍斜坡步长 [表值单位] / Ramp step this scan *)
    _fNew   : REAL;                         (* 本拍写表候选值 [表值单位] / Candidate table value *)
    _fPtPos : REAL;                         (* 目标点主轴相位位置 [度] / Target point master position *)
    _fDtSec : REAL;                         (* 扫描周期秒值，域 > eps [s] / Scan period seconds *)
    _nLo    : INT;                          (* 左邻点序号（单调验证）[点] / Left neighbor index *)
    _nHi    : INT;                          (* 右邻点序号（单调验证）[点] / Right neighbor index *)
END_VAR
VAR CONSTANT
    DL_CLT_NMIN : INT   := 2;               (* 表点数下限（边界⑥）[点] / Point count lower bound *)
    DL_CLT_NMAX : INT   := 16;              (* 表点数上限（数组容量）[点] / Point count upper bound *)
    DL_CLT_EPS  : REAL  := 1.0E-6;          (* 判零容差 [-] / Epsilon *)
END_VAR

(* —— 段 0：当拍判据派生 + 实例无条件刷新（R228A） —— *)
_fDtSec := TIME_TO_LREAL(tScan) / 1000.0;                (* 扫描周期秒化（除子常量 1000） / Scan period seconds *)
_bCfgBad := (nPts < DL_CLT_NMIN) OR (nPts > DL_CLT_NMAX) (* 点数域闸（边界⑥） / Point count gate *)
            OR (fTrimMax <= DL_CLT_EPS)                  (* 饱和上限正域闸（边界③） / Saturation gate *)
            OR (fRampRate <= DL_CLT_EPS)                 (* 斜坡率正域闸（边界④） / Ramp rate gate *)
            OR (fTol <= DL_CLT_EPS)                      (* 容差正域闸（边界①） / Tolerance gate *)
            OR (fMasterSpan <= DL_CLT_EPS)               (* 量程正域闸 / Span gate *)
            OR NOT (tScan > T#0S);                       (* 周期正域闸 / Period gate *)
rtApply(CLK := bApply);                                  (* 申请沿每拍必调 / Apply edge every scan *)
rtReset(CLK := bReset);                                  (* 复位沿每拍必调 / Reset edge every scan *)
_bFin := (fMasterPos = fMasterPos) AND ((fMasterPos - fMasterPos) = (fMasterPos - fMasterPos))   (* 主轴相位 NaN 自反 + Inf 差判闸（边界④） / Master pos NaN and Inf gate *)
         AND (fTrim = fTrim) AND ((fTrim - fTrim) = (fTrim - fTrim));   (* 修调量 NaN 自反 + Inf 差判闸 / Trim NaN and Inf gate *)
_fStep := fRampRate * _fDtSec;                           (* 斜坡步长 = 率 × 周期秒值（边界④） / Ramp step *)

(* —— 段 1：单拍量预清零（R107） —— *)
_bDoneI := FALSE;                                        (* 完成脉冲内部量预清 / Done preset *)
bTrimDone := FALSE;                                      (* 完成脉冲出口预清 / Done outlet preset *)

(* —— 段 2：复位沿处理（作用域：清故障 + 清注入状态 + 迁 eIdle，R283 逐项声明） —— *)
IF rtReset.Q THEN
    _bFault := FALSE;                                    (* 清故障锁存 / Clear fault *)
    _eCause := E_DL_CltCause.eNone;                      (* 清成因 / Clear cause *)
    _bInj := FALSE;                                      (* 清注入标志 / Clear ramping flag *)
    _fApplI := 0.0;                                      (* 清已注入量 / Clear applied *)
    fApplied := 0.0;                                     (* 清镜像出口 / Clear mirror *)
    _eState := E_DL_CltState.eIdle;                      (* 迁未使能相 / Back to idle *)
END_IF

(* —— 段 3：组态故障锁存（锁存至复位沿，R189） —— *)
IF _bCfgBad AND NOT _bFault THEN
    _bFault := TRUE;                                     (* 锁存故障位 / Latch fault *)
    _eCause := E_DL_CltCause.eCfgIllegal;                (* 成因：组态非法 / Cause illegal config *)
    _eState := E_DL_CltState.eFault;                     (* 同步迁故障相 / Migrate to fault *)
END_IF

(* —— 段 4：CASE 主状态机（ELSE 兜底迁 eFault，红线 6） —— *)
CASE _eState OF
    E_DL_CltState.eIdle:                                 (* 未使能：出口确定值 / Idle *)
        fApplied := 0.0;                                 (* 失能镜像出口清零 / Disabled mirror zero *)
        bTrimDone := FALSE;                              (* 失能完成脉冲清零 / Disabled done pulse *)
        IF bEnable AND NOT _bFault THEN
            _eState := E_DL_CltState.eRun;               (* 进入修调运行相 / Enter running *)
        END_IF
    E_DL_CltState.eRun:                                  (* 运行相：申请受理 + 相位闸斜坡注入 / Running *)
        IF NOT bEnable THEN
            _eState := E_DL_CltState.eIdle;              (* 失能回未使能（注入中止保持现状） / Back to idle *)
        ELSE
            IF rtApply.Q AND NOT _bInj AND NOT _bFault AND _bFin THEN   (* 申请受理（非注入中 + 组态在域 + 有限） / Accept request *)
                IF (nIdx >= 1) AND (nIdx <= nPts) THEN   (* 点序号域内才受理（边界⑥，申请级拒绝） / Index gate *)
                    _nIdxE := nIdx;                      (* 受理生效序号 / Effective index *)
                    _fTarget := fTrim;                   (* 目标量初值 / Target init *)
                    IF _fTarget > fTrimMax THEN
                        _fTarget := fTrimMax;            (* 正向饱和钳位（边界③） / Positive saturation *)
                    END_IF
                    IF _fTarget < (-fTrimMax) THEN
                        _fTarget := (-fTrimMax);         (* 负向饱和钳位（对称，边界③） / Negative saturation *)
                    END_IF
                    _fBase := aTable[_nIdxE];            (* 注入前基线快照（回滚锚点，边界②⑤） / Baseline snapshot *)
                    _fApplI := 0.0;                      (* 已注入量清零 / Applied zero *)
                    _bInj := TRUE;                       (* 置注入进行标志 / Ramping set *)
                END_IF
            END_IF
            IF _bInj THEN                                (* 注入进行中：相位闸 + 斜坡写表 / Ramping *)
                _fPtPos := fMasterSpan * INT_TO_REAL(_nIdxE - 1) / INT_TO_REAL(nPts - 1);   (* 目标点主轴位置（除子 = 点数-1 >= 1） / Point position *)
                IF _bFin AND (ABS(fMasterPos - _fPtPos) <= fTol) THEN   (* 相位闸：点 ± 容差窗内（边界①） / Phase gate *)
                    IF ABS(_fTarget - _fApplI) <= _fStep THEN
                        _fApplI := _fTarget;             (* 步长内直达目标 / Reach target *)
                        _bDoneI := TRUE;                 (* 完成脉冲内部置位（R187） / Done internal *)
                        _bInj := FALSE;                  (* 注入收口 / Ramping clear *)
                    ELSE
                        IF _fTarget > _fApplI THEN
                            _fApplI := _fApplI + _fStep; (* 正向斜坡步进 / Ramp up *)
                        ELSE
                            _fApplI := _fApplI - _fStep; (* 负向斜坡步进 / Ramp down *)
                        END_IF
                    END_IF
                    _fNew := _fBase + _fApplI;           (* 写表候选值 = 基线 + 已注入 / Candidate value *)
                    _nLo := _nIdxE - 1;                  (* 左邻序号 / Left neighbor *)
                    _nHi := _nIdxE + 1;                  (* 右邻序号 / Right neighbor *)
                    IF (_nLo >= 1) AND NOT (_fNew > aTable[_nLo] + DL_CLT_EPS) THEN   (* 左单调验证（容差直比） / Left monotonic check *)
                        aTable[_nIdxE] := _fBase;        (* 破坏单调回滚本点（边界②） / Rollback point *)
                        _bFault := TRUE;                 (* 锁存故障至复位沿 / Latch fault *)
                        _eCause := E_DL_CltCause.eMonotonic;   (* 成因：单调破坏 / Cause monotonic *)
                        _bInj := FALSE;                  (* 停止注入 / Stop ramping *)
                        _fApplI := 0.0;                  (* 已注入量清零 / Applied zero *)
                    ELSIF (_nHi <= nPts) AND NOT (_fNew < aTable[_nHi] - DL_CLT_EPS) THEN   (* 右单调验证 / Right monotonic check *)
                        aTable[_nIdxE] := _fBase;        (* 破坏单调回滚本点（边界②） / Rollback point *)
                        _bFault := TRUE;                 (* 锁存故障至复位沿 / Latch fault *)
                        _eCause := E_DL_CltCause.eMonotonic;   (* 成因：单调破坏 / Cause monotonic *)
                        _bInj := FALSE;                  (* 停止注入 / Stop ramping *)
                        _fApplI := 0.0;                  (* 已注入量清零 / Applied zero *)
                    ELSE
                        aTable[_nIdxE] := _fNew;         (* 单调保持：写表（随改随验） / Write table *)
                        fApplied := _fApplI;             (* 已注入量镜像出口 / Applied mirror *)
                    END_IF
                END_IF                                   (* 相位窗外：本拍不注入不写表（边界①④） *)
            END_IF
        END_IF
    E_DL_CltState.eFault:                                (* 故障相：冻结保持，仅复位沿出 / Fault *)
        ;                                                (* 锁存回放（R28） / Replay from latch *)
    ELSE                                                 (* 非法相位兜底迁安全态 / Illegal phase fallback *)
        _eState := E_DL_CltState.eFault; _bFault := TRUE;    (* 迁故障相 + 同步锁存 / To fault and latch *)
        _eCause := E_DL_CltCause.ePhaseBad;              (* 成因：非法相位 / Cause illegal phase *)
END_CASE

(* —— 段 5：出口映射（内部 _b* → 输出单拍，R187；名实双出口，R191） —— *)
bTrimDone := _bDoneI;                                    (* 完成脉冲单拍出口 / Done pulse outlet *)
bError := _bFault;                                       (* 故障标志镜像 / Fault flag mirror *)
eState := _eState;                                       (* 状态出口 / State outlet *)
eCause := _eCause;                                       (* 成因出口 / Cause outlet *)
END_FUNCTION_BLOCK

(* ---- FB_DL_CamTableOnlineBlend.st ---- *)
//==============================================================================
// 功能块：FB_DL_CamTableOnlineBlend ｜ 中文名称：凸轮表在线无缝切换（双表交叉渐变）
// 所属子库：DL_Motion ｜ 版本：v1.0.1 ｜ 日期：2026-11-23
// 兼容：CODESYS V3.5+ / TwinCAT 3 / 汇川 InoProShop（纯 IEC 61131-3 第 3 版，零方言）
// 功能描述：两张已运行的凸轮修正源（表 A / 表 B 的位置输出以引脚注入）在线
//           交叉渐变切换：切换令沿触发后，权重 w 以当前稳态值为起点、在
//           tBlend 时长内线性推进到目标值（A→B：0→1；B→A：1→0，双向可逆），
//           输出 fPosOut = (1−w)·fPosA + w·fPosB。相位连续性由权重起点连续
//           天然保证：切换瞬间 w 从稳态值起步，输出无台阶；渐变期两表输出
//           按权重交叉合成，终点严格等于目标表原样输出。
//           职责边界：本件做表级切换；表内逐点修调属 FB_DL_CamDynTrim
//           （属主已判已覆盖，互不替代）。
// 开源溯源 (Origin)：原创实现（t1-6-plcopen 表级切换语义深化，零外部源码行，
//           clean-room 独立编写；与 CamDynTrim 属主分工已在头注释声明）
// 公开接口清单：输入 bEn / bSwCmd / fPosA / fPosB / tBlend；
//               输出 fPosOut / fW / bSwitching / bSwitchDone / eState /
//               uErrCode / bValid
// 单位表：fPosA/fPosB/fPosOut[mm] / fW[1]（无量纲权重）/ tBlend[ms]
// 输入契约：fPosA/fPosB 为两表各自刷新的位置修正输出，须同一主轴位置基准；
//           tBlend 为渐变总时长，只在切换沿采纳（渐变中途改参下沿生效）。
// 输出契约：fPosOut 直接叠加主轴位置给定；fW 供上位机观察切换进度；
//           bSwitchDone 单拍完成脉冲；uErrCode 信息级不锁存；
//           bValid = FALSE 拍输出冻结为上一拍有效合成快照（首拍即非有限、
//           无快照时哨兵 0.0）。
// 错误码表：16#0004_08D0 信息级（切换时长非法拒绝触发、位置源非有限安全侧
//           冻结输出，不置 bError）/ 16#0004_08D1 预留禁用（不得挪用）
// 状态机：E_DL_CamBlendState（本文件唯一定义，全库唯一属主）：
//           eActive = 0 / eBlending = 10
// 边界行为：① tBlend <= 0 或非有限 → 拒绝触发 + 信息码，保持当前表原样；
//           ② 位置源非有限 → 输出冻结上一拍有效快照 _fPosOutLast 直通
//             fPosOut，非法输入不参与任何算术；无快照（首拍即非有限）哨兵
//             0.0 + bValid := FALSE（安全侧，R73 返修）；
//           ③ 权重起点/终点在切换沿单拍锁存，渐变期内不刷新（连续性关键）；
//           ④ w 全程钳 0..1，时长换算用 TIME_TO_LREAL（库内已证可编译口径，R397 弃用 TIME_TO_DWORD 非标准扩展）；
//           ⑤ CASE 带 ELSE 非法态兜底回 eActive；
//           ⑥ TON/R_TRIG 每拍无条件刷新（不入分支，红线 R7）；
//           ⑦ 渐变期内重复切换令被抑制（信息级留痕不打断权重窗，
//             R90 复用码）。
// 修订历史：v1.0.0 2026-11-23 首版（R73 派单 · 批 1 · 序 2）
//           v1.0.1 2026-11-23 R73 返修：非有限防御分支改冻结上一拍有效输出
//           快照（新增 _fPosOutLast / _bOutValid，无条件段统一滚存），非法
//           输入不再参与合成算术，NaN/Inf 不直穿输出。
//==============================================================================

(*------------------------------------------------------------------------------
 * 枚举: E_DL_CamBlendState（归属本功能块，同文件发布，全库唯一属主）
 * 含义: 双表切换相位，成员与 CASE 标签双向完备。
 *-----------------------------------------------------------------------------*)
TYPE E_DL_CamBlendState :
(
    eActive   := 0,    // 稳态：按当前权重直接输出 / Steady state, output by the current weight
    eBlending := 10    // 渐变中：权重向目标值线性推进 / Blending, weight advancing toward the target
);
END_TYPE

(*==============================================================================
 * 功能块: FB_DL_CamTableOnlineBlend
 * 调用约定: 每个扫描周期无条件调用一次；实例状态全部驻留于私有变量。
 * 调用示例: camBlend(bEn := TRUE, bSwCmd := bSwSelB,
 *                    fPosA := camTableA.fCorr, fPosB := camTableB.fCorr,
 *                    tBlend := T#2S);
 *          两表各自独立刷新修正输出后经引脚注入；合成输出
 *          camBlend.fPosOut 直接叠加到主轴位置给定上。
 * 组装说明: ① 两张凸轮表的逐点修调由各自表实例承担（CamDynTrim 属主），
 *             本件只消费两表的输出引脚，不触碰表数据本体；
 *           ② bSwCmd 双向触发：当前权重 < 0.5 判向 B 表渐变，反之判向
 *             A 表，回切无需反向专用引脚；
 *           ③ 切换期间禁止上层同时改 tBlend（时长闸只在触发沿生效，
 *             渐变中途改参将被下一次沿才采纳）；
 *           ④ 位置源非有限时输出冻结上一有效权重合成值并拉低 bValid，
 *             上层应据 bValid 门控下游位置给定的采纳。
 *==============================================================================*)
FUNCTION_BLOCK FB_DL_CamTableOnlineBlend
VAR_INPUT
    bEn      : BOOL := FALSE;          // 使能（FALSE 冻结输出并回稳态）/ Enable, FALSE freezes and returns to steady
    bSwCmd   : BOOL := FALSE;          // 切换令沿：双向，触发即向目标表渐变 / Switch command edge, bidirectional, trigger blends toward the target table
    fPosA    : LREAL := 0.0;           // 表 A 位置修正输出 [mm]，引脚注入 / Table A position output [mm], injected via the pin
    fPosB    : LREAL := 0.0;           // 表 B 位置修正输出 [mm]，引脚注入 / Table B position output [mm], injected via the pin
    tBlend   : TIME  := T#1S;          // 渐变时长 [ms]，权窗推进总时长 / Blend duration [ms], total weight window
END_VAR
VAR_OUTPUT
    fPosOut  : LREAL;                  // 交叉合成位置输出 [mm] / Crossfaded position output [mm]
    fW       : LREAL;                  // 当前权重 w [1]，0 = 全 A / 1 = 全 B / Current blend weight [1]
    bSwitching: BOOL;                  // TRUE = 渐变进行中 / TRUE = blending in progress
    bSwitchDone: BOOL;                 // 单拍切换完成脉冲 / Single-scan switch-done pulse
    eState   : E_DL_CamBlendState;     // 切换当前相位 / Current blend phase
    uErrCode : UDINT;                  // 信息级码，0 = 无信息 / Info-level code, 0 = none
    bValid   : BOOL;                   // 输出有效标志 / Outputs usable flag
END_VAR
VAR
    tonBlend : TON;                    // 渐变权窗定时器，每拍无条件刷新 / Blend weight timer, refreshed every scan
    trigSw   : R_TRIG;                 // 切换令沿检测，每拍无条件刷新 / Switch command edge, refreshed every scan
    fWStart  : LREAL;                  // 渐变起点权重 [1]，切换沿锁存 / Start weight [1], latched at the switch edge
    fWEnd    : LREAL;                  // 渐变终点权重 [1]，切换沿锁存 / End weight [1], latched at the switch edge
    _bDone   : BOOL;                   // 完成脉冲内部暂存（统一出口映射） / Done stage internal, mapped at the unified outlet
    _fPosOutLast : LREAL;              // 上一拍有效合成输出快照 [mm]，非有限拍冻结源 / Last valid output snapshot [mm], freeze source on non-finite scans
    _bOutValid   : BOOL;               // 快照有效声明（首个有效拍后置位）/ Snapshot validity flag, set after the first valid scan
END_VAR
VAR CONSTANT
    DL_CB_EPS  : LREAL := 1.0E-9;      // 浮点容差 / Float tolerance
    DL_CB_INF  : LREAL := 1.7976931348623157E308; // LREAL 幅值上限 / LREAL magnitude ceiling
    DL_CB_WMIN : LREAL := 0.0;         // 权重下界 [1]，全 A 表 / Weight floor [1], table A only
    DL_CB_WMAX : LREAL := 1.0;         // 权重上界 [1]，全 B 表 / Weight ceiling [1], table B only
END_VAR

// ---- 段 1｜定时/沿实例无条件刷新 + 单拍脉冲出口预清（红线 R7 + 两段式）----
tonBlend(IN := (eState = E_DL_CamBlendState.eBlending), PT := tBlend); // 权窗计时按态断输入 / Weight timer input per state
trigSw(CLK := bSwCmd);                 // 切换令沿每拍刷新 / Switch edge refreshed unconditionally
_bDone      := FALSE;                  // 完成脉冲暂存先清零 / Done stage preset FALSE
bSwitching  := FALSE;                  // 渐变声明默认 FALSE / Switching flag preset FALSE
bSwitchDone := FALSE;                  // 完成脉冲默认 FALSE（相内重置位）/ Done pulse preset FALSE
uErrCode    := 16#0000_0000;           // 信息码每拍重算（信息级不锁存）/ Info code recomputed, info level never latched
bValid      := TRUE;                   // 可用标志默认 TRUE（防御段可改写）/ Usable flag preset TRUE, defense may overwrite

// ---- 段 2｜输入防御：位置源或时长非有限 → 输出冻结 + 安全侧回稳态 ----
IF (fPosA <> fPosA) OR (ABS(fPosA) > DL_CB_INF)
   OR (fPosB <> fPosB) OR (ABS(fPosB) > DL_CB_INF) THEN
    uErrCode := 16#0004_08D0;          // 信息级：位置源非有限 / Info: non-finite position source
    bValid   := FALSE;                 // 输出不可用 / Outputs unusable
    IF eState <> E_DL_CamBlendState.eActive THEN
        eState := E_DL_CamBlendState.eActive; // 渐变中止回稳态（权重保持当前值）/ Blending aborted, weight held
    END_IF
    IF _bOutValid THEN                 // 已有有效快照 → 冻结直通 / Snapshot available, freeze through
        fPosOut := _fPosOutLast;       // 冻结上一拍有效输出（非法输入不参与算术）/ Freeze the last valid output, invalid input never enters arithmetic
    ELSE
        fPosOut := 0.0;                // 首拍即非有限无快照：哨兵 0.0 / Non-finite on the first scan, sentinel zero
    END_IF
    RETURN;                            // 结构早退 / early exit
END_IF

// ---- 段 3｜状态机（CASE 带 ELSE；权重推进除法先过时长闸）----
CASE eState OF
    E_DL_CamBlendState.eActive:        // 稳态相：按当前权重合成输出
        fPosOut := fW * fPosB + (1.0 - fW) * fPosA; // 交叉合成 [mm] / Crossfade blend [mm]
        IF bEn AND trigSw.Q AND (tBlend > T#0MS) THEN
            IF fW < (0.5 + DL_CB_EPS) THEN // 距 B 更近判目标（中点判决）/ Target table by midpoint decision
                fWStart := fW;             // 起点权重锁存（连续性关键）/ Start weight latched, the continuity key
                fWEnd   := DL_CB_WMAX;     // 目标权重 1（B 表）/ Target weight 1, table B
            ELSE
                fWStart := fW;             // 起点权重锁存 / Start weight latched
                fWEnd   := DL_CB_WMIN;     // 目标权重 0（A 表）/ Target weight 0, table A
            END_IF
            eState := E_DL_CamBlendState.eBlending; // 进入渐变相 / Enter the blending phase
        END_IF

    E_DL_CamBlendState.eBlending:      // 渐变相：权重向目标值线性推进，输出相位连续
        bSwitching := TRUE;            // 渐变进行中声明 / Blending declared
        IF trigSw.Q THEN               // 渐变期内重复切换令抑制（信息级留痕，不打断权重窗）/ Repeated command suppressed, info trace
            uErrCode := 16#0004_08D0;  // 信息级：切换令被抑制（复用码 R90）/ Info: command suppressed, code reused per R90
        END_IF
        IF tBlend > T#0MS THEN         // 时长闸（防除零前置，双保险复检）/ Duration gate, defense in depth
            fW := fWStart + (fWEnd - fWStart)
                  * TIME_TO_LREAL(tonBlend.ET)
                  / TIME_TO_LREAL(tBlend);      // 权重线性推进 [1] / Linear weight advance [1]
        END_IF
        fW := MIN(MAX(fW, DL_CB_WMIN), DL_CB_WMAX); // 权重双侧钳位 / Two-sided weight clamp
        fPosOut := fW * fPosB + (1.0 - fW) * fPosA; // 相位连续合成 [mm] / Phase-continuous blend [mm]
        IF tonBlend.Q THEN
            fW     := fWEnd;           // 权窗到顶强制终点值（防尾差）/ Force the end weight at window end
            eState := E_DL_CamBlendState.eActive; // 渐变完成回稳态 / Blending complete, back to steady
            _bDone := TRUE;            // 完成脉冲内部置位（出口统一映射） / Done stage set for the outlet
        END_IF

    ELSE                               // 非法状态兜底（R21：CASE 必带 ELSE）
        eState  := E_DL_CamBlendState.eActive; // 拦截非法值回稳态 / Catch illegal value back to steady
        fW      := DL_CB_WMIN;         // 权重回 0（A 表侧安全）/ Weight back to 0, table A side
        fPosOut := fPosA;              // 输出回 A 表原样 / Output back to table A as-is
END_CASE

// ---- 段 4｜统一出口：完成脉冲单拍映射 + 撤使能兜底 ----
IF NOT bEn THEN                        // 撤使能兜底（门控挂状态量，非单拍标志）
    IF eState <> E_DL_CamBlendState.eActive THEN
        eState  := E_DL_CamBlendState.eActive; // 回稳态 / Back to steady state
        fW      := DL_CB_WMIN;         // 权重回 0 / Weight back to zero
    END_IF
    fPosOut := fPosA;                  // 撤使能输出回 A 表原样 / Disabled output back to table A
END_IF
bSwitchDone := _bDone;                 // 完成脉冲本拍有效（两段式出口）/ Done pulse valid this scan
_fPosOutLast := fPosOut;               // 快照滚存（到达此处输入必已过有限闸）/ Snapshot rolled forward, the finite gate already passed
_bOutValid   := TRUE;                  // 快照有效声明 / Snapshot declared valid
END_FUNCTION_BLOCK

(* ---- FB_DL_CircInterp2Axis.st ---- *)
(*
  组件名 Component   : FB_DL_CircInterp2Axis
  子库 Sublibrary    : DL_Motion
  版本 Version       : 1.0.0
  兼容性 Platform    : CODESYS 3.5 / TwinCAT 3 / 汇川 InoProShop / Machine Expert（仅 Standard.library）
  功能 Function      : 两轴圆弧插补（与 FB_DL_LineInterp2Axis 同线直角补口）：
                       1) 双模式几何解算：圆心模式（半径由起点到圆心距实测，终点距圆心
                       超容差判组态非法）/ 半径模式（由起终点弦长与半径反解圆心，CW/CCW
                       定唯一解，弦长 > 2R 判组态非法）；
                       2) 弓高误差弦长分段：每拍角步长 = 进给/半径 与 弦长上限角步长
                       取小（弦长上限由弓高误差限反解，半径/进给除法前置域闸）；
                       3) 象限跨越判据：本拍与上拍象限号不同 → bQuadCross 单拍脉冲；
                       4) 终点判定：剩余弧角 <= 步长 → 落终点，eDone 驻留。
  边界 Boundary      : ① 本件只出两轴位置设定点，不接管轴使能与物理 IO；
                       ② 角度归一化循环带守卫计数器（上限 8 次，超限判几何非法）；
                       ③ 反三角经 FC_DL_Atan2Ex 唯一属主（DL_MathData），本件零重写；
                       ④ 非有限值（NaN 自反 + 无穷差值自减）判非法锁存，出点冻结；
                       ⑤ 故障锁存解除唯一路径 = bReset 上升沿（输入引脚，恒可达）；
                       ⑥ 无全局变量引用、无外部变量声明、无物理地址寻址。
  依赖 Depends       : FC_DL_Atan2Ex（DL_MathData，按 registry 实名）；Standard.library（R_TRIG）
  溯源 Origin        : 道莅自研 clean-room（参考 t1-8-github motion 线分类与参数域，
                       零代码行复制；圆弧参数化与弓高分段为公开几何语义）
  码位 Code          : 16#04_0_AC
  码表 Error codes（Motion 格 04_0_AC，单轨：故障 0x02AC / 信息 0x01AC）:
    16#0004_02AC 故障级：几何解算非法（弦长 > 2R / 终点半径超容差 / 进给或弓高限
                 非法 / 输入非有限 / 归一化守卫超限），锁存至 bReset 上升沿
    16#0004_01AC 信息级：象限跨越脉冲沿（bQuadCross 置位拍）
  修订历史 Revision  :
    2026-11-19  v1.0.0  R44 首版（批次 2 · 序号 9）
*)

TYPE E_DL_CiaState :
(
    eIdle   := 0,   // 空闲：等启动沿 / Idle, waiting start edge
    eGeom   := 10,  // 几何：单拍解算圆心/半径/弧角 / Geometry, one-pass solve
    eRun    := 20,  // 插补：逐拍步进出点 / Interpolating, per-scan stepping
    eDone   := 30,  // 完成：落终点驻留 / Done, at end point
    eFault  := 90   // 故障：几何/输入锁存 / Fault, latched
);
END_TYPE

FUNCTION_BLOCK FB_DL_CircInterp2Axis
VAR_INPUT
    bStartCmd    : BOOL;                   // 启动指令（上升沿承载）[-] / Start command edge
    bReset       : BOOL;                   // 上升沿清故障锁存 [-] / Reset edge
    fStartXMm    : REAL;                   // 起点坐标 X [mm] / Start point X
    fStartYMm    : REAL;                   // 起点坐标 Y [mm] / Start point Y
    fEndXMm      : REAL;                   // 终点坐标 X [mm] / End point X
    fEndYMm      : REAL;                   // 终点坐标 Y [mm] / End point Y
    bUseRadius   : BOOL;                   // 模式：TRUE = 半径模式 / Mode, TRUE = radius mode
    fCenterXMm   : REAL;                   // 圆心坐标 X（圆心模式）[mm] / Center X
    fCenterYMm   : REAL;                   // 圆心坐标 Y（圆心模式）[mm] / Center Y
    fRadiusMm    : REAL;                   // 半径（半径模式）[mm] / Radius
    bCwDir       : BOOL;                   // 方向：TRUE = 顺时针 [-] / Direction, TRUE = CW
    fFeedMmS     : REAL := 50.0;           // 合成进给速度 [mm/s] / Feed velocity
    fSagittaMaxMm: REAL := 0.01;           // 弓高误差限 [mm] / Sagitta error limit
    fRadTolMm    : REAL := 0.01;           // 终点半径容差 [mm] / End radius tolerance
    tCycle       : TIME := T#10MS;         // 扫描周期 [毫秒] / Scan cycle time
END_VAR
VAR_OUTPUT
    fPosXMm      : REAL;                   // 位置设定点 X [mm] / Position setpoint X
    fPosYMm      : REAL;                   // 位置设定点 Y [mm] / Position setpoint Y
    bBusy        : BOOL;                   // 插补进行中电平 [-] / Interpolation busy
    bDone        : BOOL;                   // 到达终点电平 [-] / End-point reached level
    bQuadCross   : BOOL;                   // 象限跨越单拍脉冲 [-] / Quadrant crossing pulse
    fArcLenMm    : REAL;                   // 解算弧长 [mm] / Computed arc length
    eState       : E_DL_CiaState;          // 状态出口，段尾单点映射 / State outlet
    bError       : BOOL;                   // 故障锁存标志 [-] / Fault latch flag
    uErrId       : UDINT;                  // 事件码，0 = 无事件 / Event code
END_VAR
VAR
    rtReset : R_TRIG;                      // 复位沿实例，段 0 无条件刷新 / Reset edge
    rtStart : R_TRIG;                      // 启动沿实例，段 0 无条件刷新 / Start edge
    _eState : E_DL_CiaState := E_DL_CiaState.eIdle;    // 内部相位（CASE 唯一写入目标）/ Internal phase
    _fCtrXMm: REAL;                        // 解算圆心 X [mm] / Solved center X
    _fCtrYMm: REAL;                        // 解算圆心 Y [mm] / Solved center Y
    _fRadMm : REAL;                        // 解算半径 [mm] / Solved radius
    _fAng0  : REAL;                        // 起点角 [弧度] / Start angle
    _fAng1  : REAL;                        // 终点角 [弧度] / End angle
    _fSweep : REAL;                        // 弧角绝对扫角 [弧度] / Absolute sweep
    _fAngCur: REAL;                        // 当前角 [弧度] / Current angle
    _fDAng  : REAL;                        // 每拍角步长 [弧度] / Angular step per scan
    _nQuadPrev: DINT;                      // 上拍象限号 [-] / Previous quadrant
    _nQuadCur : DINT;                      // 本拍象限号 [-] / Current quadrant
    _bFault : BOOL;                        // 故障锁存位（锁存量） / Latched fault bit
    _uFault : UDINT;                       // 故障码锁存（锁存量） / Latched fault code
    _bCfgBad: BOOL;                        // 组态非法当拍量 [-] / Config illegal flag
    _bNonFin: BOOL;                        // 输入非有限当拍量 [-] / Non-finite input flag
    _bValid : BOOL;                        // Atan2Ex 属主返回有效标志（两调用与集） / Atan2 validity flag
    _bVal0  : BOOL;                        // 起点角属主有效标志 [-] / Start angle validity
    _bVal1  : BOOL;                        // 终点角属主有效标志 [-] / End angle validity
    fDxGeom : LREAL;                       // 几何解算弦向量 X [mm] / Geometry chord vector X
    fDyGeom : LREAL;                       // 几何解算弦向量 Y [mm] / Geometry chord vector Y
    fChordGeom : LREAL;                    // 几何解算弦长 [mm] / Geometry chord length
    fHGeom  : LREAL;                       // 圆心偏距 [mm] / Center offset distance
    fAng0Geom : LREAL;                     // 起点角属主返回值 [弧度] / Start angle owner result
    fAng1Geom : LREAL;                     // 终点角属主返回值 [弧度] / End angle owner result
    fSweepGeom: LREAL;                     // 扫角归一化中间量 [弧度] / Sweep normalization temp
    _nNormGuard: DINT;                     // 归一化守卫计数 [次] / Normalization guard counter
    fStepFeed : LREAL;                     // 进给角步长 [弧度] / Feed angular step
    fChordMax : LREAL;                     // 弓高弦长上限 [mm] / Sagitta chord ceiling
    fStepGeom : LREAL;                     // 弦长上限角步长 [弧度] / Chord-ceiling angular step
    fRemainGeom: LREAL;                    // 剩余扫角 [弧度] / Remaining sweep
END_VAR
VAR CONSTANT
    DL_TWO_PI  : REAL := 6.283185307;      // 全周角 [弧度] / Full turn angle
    DL_HALF_PI : REAL := 1.570796327;      // 直角 [弧度] / Quarter turn angle
    DL_TWO     : REAL := 2.0;              // 二常量 [无量纲] / Two constant
    DL_EPS     : REAL := 1.0E-6;           // 几何退化判据 [mm] / Degenerate geometry tolerance
    DL_NORM_GUARD: DINT := 8;              // 角度归一化守卫上限 [次] / Normalization guard limit
    DL_ABS_MAX : REAL := 1.0E30;           // 有限值判定上界 [mm] / Finite bound
    DL_ZERO    : REAL := 0.0;              // 零常量 [mm] / Zero constant
    DL_MS_PER_S: REAL := 1000.0;           // 毫秒 → 秒换算系数 [毫秒/秒] / Milliseconds per second
END_VAR

(* —— 段 0｜沿实例每拍无条件刷新（禁置于 IF/CASE 内） —— *)
rtReset(CLK := bReset);
rtStart(CLK := bStartCmd);

(* —— 段 1｜瞬时量预清零（锁存量 _bFault/_uFault/bDone/几何量不入清单） —— *)
uErrId     := 16#0000_0000;
bQuadCross := FALSE;                     // 跨越脉冲单拍量，每拍清零
_bCfgBad   := FALSE;
_bNonFin   := FALSE;
_bValid    := TRUE;

(* —— 段 2｜复位沿：故障一次性清干净，相位回空闲 —— *)
IF rtReset.Q THEN
    _bFault := FALSE;
    _uFault := 16#0000_0000;
    bDone   := FALSE;
    _eState := E_DL_CiaState.eIdle;
END_IF

(* —— 段 3｜公共组态闸与非有限判据（覆盖全部参与换算引脚） —— *)
IF (fFeedMmS <= DL_ZERO) OR (fSagittaMaxMm <= DL_ZERO) OR (fRadTolMm <= DL_ZERO)
   OR (tCycle = T#0S) THEN
    _bCfgBad := TRUE;
END_IF
IF (fStartXMm <> fStartXMm) OR ((fStartXMm - fStartXMm) <> DL_ZERO)
   OR (fStartYMm <> fStartYMm) OR ((fStartYMm - fStartYMm) <> DL_ZERO)
   OR (fEndXMm <> fEndXMm) OR ((fEndXMm - fEndXMm) <> DL_ZERO)
   OR (fEndYMm <> fEndYMm) OR ((fEndYMm - fEndYMm) <> DL_ZERO) THEN
    _bNonFin := TRUE;
END_IF

(* —— 段 4｜主状态机：五态全覆盖 + ELSE 兜底 —— *)
CASE _eState OF

E_DL_CiaState.eIdle:
    bBusy := FALSE;
    IF rtStart.Q AND (NOT _bFault) AND (NOT _bCfgBad) AND (NOT _bNonFin) THEN
        fPosXMm := fStartXMm;            // 出点先落起点
        fPosYMm := fStartYMm;
        bDone   := FALSE;
        _eState := E_DL_CiaState.eGeom;
    ELSIF rtStart.Q AND (_bFault OR _bCfgBad OR _bNonFin) THEN
        _bFault := TRUE;                 // 带病启动拒绝
        _uFault := 16#0004_02AC;
        bError  := TRUE;
        _eState := E_DL_CiaState.eFault;
    END_IF

E_DL_CiaState.eGeom:
    (* 单拍几何解算：圆心 / 半径 / 起终角 / 扫角 *)
    IF _bNonFin THEN
        _bFault := TRUE;
        _uFault := 16#0004_02AC;
        bError  := TRUE;
        _eState := E_DL_CiaState.eFault;
    ELSE
        IF bUseRadius THEN
            (* 半径模式：弦长反解圆心（CW/CCW 定唯一解），弦长 > 2R 判非法 *)
            _fRadMm := ABS(fRadiusMm);
            IF _fRadMm <= DL_EPS THEN
                _bFault := TRUE;
                _uFault := 16#0004_02AC;
                bError  := TRUE;
                _eState := E_DL_CiaState.eFault;
            ELSE
                fDxGeom := fEndXMm - fStartXMm;          // 弦向量 X
                fDyGeom := fEndYMm - fStartYMm;          // 弦向量 Y
                fChordGeom := SQRT(fDxGeom * fDxGeom + fDyGeom * fDyGeom);
                IF fChordGeom <= DL_EPS THEN
                    _bFault := TRUE;     // 起终点重合：圆弧退化
                    _uFault := 16#0004_02AC;
                    bError  := TRUE;
                    _eState := E_DL_CiaState.eFault;
                ELSIF fChordGeom > (DL_TWO * _fRadMm) THEN
                    _bFault := TRUE;     // 弦长超直径：无解
                    _uFault := 16#0004_02AC;
                    bError  := TRUE;
                    _eState := E_DL_CiaState.eFault;
                ELSE
                    fHGeom := SQRT(MAX(_fRadMm * _fRadMm - (fChordGeom * fChordGeom) / (DL_TWO * DL_TWO), DL_ZERO));
                    _fCtrXMm := (fStartXMm + fEndXMm) / DL_TWO;
                    _fCtrYMm := (fStartYMm + fEndYMm) / DL_TWO;
                    IF bCwDir THEN
                        _fCtrXMm := _fCtrXMm + (fDyGeom / fChordGeom) * fHGeom;
                        _fCtrYMm := _fCtrYMm - (fDxGeom / fChordGeom) * fHGeom;
                    ELSE
                        _fCtrXMm := _fCtrXMm - (fDyGeom / fChordGeom) * fHGeom;
                        _fCtrYMm := _fCtrYMm + (fDxGeom / fChordGeom) * fHGeom;
                    END_IF
                    _eState := E_DL_CiaState.eRun;
                END_IF
            END_IF
        ELSE
            (* 圆心模式：半径由起点实测，终点半径超容差判非法 *)
            _fCtrXMm := fCenterXMm;
            _fCtrYMm := fCenterYMm;
            fDxGeom := fStartXMm - _fCtrXMm;
            fDyGeom := fStartYMm - _fCtrYMm;
            _fRadMm := SQRT(fDxGeom * fDxGeom + fDyGeom * fDyGeom);
            fDxGeom := fEndXMm - _fCtrXMm;
            fDyGeom := fEndYMm - _fCtrYMm;
            fChordGeom := SQRT(fDxGeom * fDxGeom + fDyGeom * fDyGeom);
            IF _fRadMm <= DL_EPS THEN
                _bFault := TRUE;         // 起点与圆心重合
                _uFault := 16#0004_02AC;
                bError  := TRUE;
                _eState := E_DL_CiaState.eFault;
            ELSIF ABS(fChordGeom - _fRadMm) > fRadTolMm THEN
                _bFault := TRUE;         // 终点半径与起点半径超容差
                _uFault := 16#0004_02AC;
                bError  := TRUE;
                _eState := E_DL_CiaState.eFault;
            ELSE
                _eState := E_DL_CiaState.eRun;
            END_IF
        END_IF
        IF _eState = E_DL_CiaState.eRun THEN
            (* 起终角经 Atan2Ex 唯一属主（返回弧度），属主无效即判故障 *)
            fAng0Geom := FC_DL_Atan2Ex(lrY := fStartYMm - _fCtrYMm, lrX := fStartXMm - _fCtrXMm,
                                       bValid => _bVal0);
            fAng1Geom := FC_DL_Atan2Ex(lrY := fEndYMm - _fCtrYMm, lrX := fEndXMm - _fCtrXMm,
                                       bValid => _bVal1);
            _bValid := _bVal0 AND _bVal1;
            IF NOT _bValid THEN
                _bFault := TRUE;
                _uFault := 16#0004_02AC;
                bError  := TRUE;
                _eState := E_DL_CiaState.eFault;
            ELSE
                IF bCwDir THEN
                    fSweepGeom := fAng0Geom - fAng1Geom;
                ELSE
                    fSweepGeom := fAng1Geom - fAng0Geom;
                END_IF
                _nNormGuard := 0;
                WHILE (fSweepGeom < DL_ZERO) AND (_nNormGuard < DL_NORM_GUARD) DO
                    fSweepGeom := fSweepGeom + DL_TWO_PI;    // 负角加全周归一
                    _nNormGuard := _nNormGuard + 1;
                END_WHILE;
                _nNormGuard := 0;
                WHILE (fSweepGeom >= DL_TWO_PI) AND (_nNormGuard < DL_NORM_GUARD) DO
                    fSweepGeom := fSweepGeom - DL_TWO_PI;    // 超全周减全周归一
                    _nNormGuard := _nNormGuard + 1;
                END_WHILE;
                IF (_nNormGuard >= DL_NORM_GUARD) OR (fSweepGeom <= DL_EPS) THEN
                    _bFault := TRUE;     // 归一化守卫超限或扫角退化
                    _uFault := 16#0004_02AC;
                    bError  := TRUE;
                    _eState := E_DL_CiaState.eFault;
                ELSE
                    _fSweep  := LREAL_TO_REAL(fSweepGeom);
                    _fAng0   := LREAL_TO_REAL(fAng0Geom);
                    _fAngCur := _fAng0;
                    fArcLenMm := _fSweep * _fRadMm;
                    (* 每拍角步长：进给步长与弓高弦长上限步长取小（除数均已过域闸） *)
                    fStepFeed := fFeedMmS * TIME_TO_REAL(tCycle) / DL_MS_PER_S / _fRadMm;
                    fChordMax := DL_TWO * SQRT(DL_TWO * _fRadMm * fSagittaMaxMm
                                 - fSagittaMaxMm * fSagittaMaxMm);
                    fStepGeom := fChordMax / _fRadMm;
                    _fDAng := LREAL_TO_REAL(MIN(fStepFeed, fStepGeom));
                    _nQuadPrev := -1;    // 象限号初始化为哨兵
                    bBusy := TRUE;
                END_IF
            END_IF
        END_IF
    END_IF

E_DL_CiaState.eRun:
    bBusy := TRUE;
    IF bCwDir THEN
        _fAngCur := _fAngCur - _fDAng;
    ELSE
        _fAngCur := _fAngCur + _fDAng;
    END_IF
    (* 象限号判据：cos/sin 符号四象限编码（0..3），本上拍不同即跨越 *)
    IF COS(_fAngCur) >= DL_ZERO THEN
        IF SIN(_fAngCur) >= DL_ZERO THEN
            _nQuadCur := 0;              // 第一象限
        ELSE
            _nQuadCur := 3;              // 第四象限
        END_IF
    ELSE
        IF SIN(_fAngCur) >= DL_ZERO THEN
            _nQuadCur := 1;              // 第二象限
        ELSE
            _nQuadCur := 2;              // 第三象限
        END_IF
    END_IF
    IF (_nQuadPrev >= 0) AND (_nQuadCur <> _nQuadPrev) THEN
        bQuadCross := TRUE;              // 象限跨越脉冲（单拍）
        uErrId := 16#0004_01AC;          // 信息级：象限跨越沿
    END_IF
    _nQuadPrev := _nQuadCur;
    (* 出点由圆心 + 半径 × 当前角三角合成（正解三角为 Standard.library 标准函数） *)
    fPosXMm := _fCtrXMm + COS(_fAngCur) * _fRadMm;
    fPosYMm := _fCtrYMm + SIN(_fAngCur) * _fRadMm;
    (* 终点判定：剩余扫角耗尽 → 落终点驻留 *)
    fRemainGeom := ABS(_fAngCur - _fAng0);
    IF fRemainGeom >= (_fSweep - _fDAng) THEN
        fPosXMm := fEndXMm;
        fPosYMm := fEndYMm;
        bBusy := FALSE;
        bDone := TRUE;
        _eState := E_DL_CiaState.eDone;
    END_IF

E_DL_CiaState.eDone:
    bDone := TRUE;
    bBusy := FALSE;
    IF NOT bStartCmd THEN
        _eState := E_DL_CiaState.eIdle;  // 启动指令撤销：回空闲
    END_IF

E_DL_CiaState.eFault:
    bBusy := FALSE;
    bError := TRUE;
    ;                                    // 故障相驻留：出点冻结，只认复位沿（段 2 迁出）

ELSE
    _bFault := TRUE;                     // 兜底：非法相位锁存
    _uFault := 16#0004_02AC;
    bError  := TRUE;
    _eState := E_DL_CiaState.eFault;
END_CASE

(* —— 段 5｜状态出口单点映射 —— *)
eState := _eState;
END_FUNCTION_BLOCK

(* ---- FB_DL_ContourCrossCouple.st ---- *)
(*==============================================================================
 * 组件名称 (Component)  : FB_DL_ContourCrossCouple
 * 所属子库 (Sublibrary) : DL_Motion
 * 当前版本 (Version)    : 1.0.1
 * 兼容性   (Platform)   : CODESYS 3.5+ / TwinCAT 3 / 汇川 InoProShop / 施耐德 Machine Expert
 *                         仅依赖 Standard.library（ABS / SQRT / MAX），零厂商私有库
 * 功能描述 (Function)   : 双轴轮廓交叉耦合控制（闭环修调侧）：由两轴跟随误差合成轮廓误差
 *                           fEc = (fErrX×fDirX + fErrY×fDirY) / SQRT(fDirX²+fDirY²)
 *                         （fDirX/fDirY 为轨迹方向单位向量分量，组态输入），再把轮廓误差
 *                         垂直分量还给弱轴：
 *                           fTrimY = +fKc × fEc × fDirX
 *                           fTrimX = -fKc × fEc × fDirY
 *                         输出限幅 ±fTrimMaxMm；bEnable 退出时修调斜坡归零（禁突跳）；
 *                         使能期输出同样按 fRampMmS 斜率逼近目标值（换段方向向量突变
 *                         不产生阶跃）。
 * 接口     (Interface)  : 输入 fErrX/fErrY 两轴跟随误差（mm）、fDirX/fDirY 轨迹方向向量
 *                         分量（无量纲）、fKc 交叉耦合增益（0~1）、fTrimMaxMm 修调限幅
 *                         （mm）、fRampMmS 修调变化率限（mm/s）、fCycle 扫描周期（s，
 *                         <=0 用缺省）、bEnable 使能、bReset 复位；输出 fTrimX/fTrimY
 *                         修调注入（mm）、bNoDir 方向向量退化、bError 故障标志。
 * 边界     (Boundary)   : ① **属主边界（写死）：本件只算修调注入量，不写轴位置指令、
 *                         不接管插补器**；注入点由上层叠加到从轴位置设定。
 *                         ② 方向向量模 < 1E-6 → 直通零修调并置 bNoDir（R28 防零，不开方
 *                         负数/除零）。
 *                         ③ 非有限误差冻结当拍斜坡目标（保持逼近上一目标，R245）。
 *                         ④ 斜坡归零：bEnable=FALSE 时目标=0，输出按 fRampMmS×fCycle 向 0
 *                         收敛（R191 名实双出口声明：未使能期修调**斜坡归零而非保持**）。
 *                         ⑤ 组态闸：fKc<0 或 >1、fTrimMaxMm<=0、fRampMmS<=0 → 锁存
 *                         bError，输出强制归零，解除沿 = bReset 上升沿。
 *                         ⑥ 零全局耦合（无 GVL / VAR_EXTERNAL / 物理地址）。
 * 分工声明 (Scope)      : 与 `FB_DL_GantrySkewMonitor` 分工：闭环修调（本件）≠ 偏差监视
 *                         （那件）；与 `FB_DL_LoadShareDroop` 分工：轮廓误差耦合 ≠ 负载
 *                         调差。
 * 来源标签 (Source Tag) : T1-6 ◐（PLCopen MC 语义只借轮廓误差定义口径，交叉耦合法则为
 *                         公开控制理论定义 clean-room）
 * 码表     (Codes)      : 本件不占用任何全局数字码位。出口为 LREAL 修调组 + BOOL 组；
 *                         数字码位待主控收口阶段统一派号。
 * 红线自检 (Redline)    : R1 ✓ 零 GVL/VAR_EXTERNAL ｜ R2 ✓ 零 %I/%Q/%M ｜ R3 ✓ 纯 IEC 61131-3
 *                         R4 ✓ 向量模防零 + 周期缺省闸 + 非有限冻结 + 限幅 ｜ R5 ✓ 声明逐行同行双语注释
 *                         R6 N/A（无状态机） ｜ R7 ✓ 一 R_TRIG 段 0 无条件刷新
 * 修订历史 (Revision)   : 2026-11-20  v1.0.1  R50 返修 R4：fDirX/fDirY 非有限
 *                         判据补 Inf 判（差自减 (x−x) <> 0），与 fErrX/fErrY
 *                         两侧口径一致（R79 双判对齐）；行为变更：方向向量
 *                         ±Inf 现判非有限冻结（原放行），验收向量同步补组。
 *                         2026-11-20  v1.0.0  R48 首版（批次 4 · 序号 16）
 *                         验收向量：X 误差主导 + 方向沿 X → fTrimY 修调、fTrimX 近零；
 *                         方向模 0 → bNoDir 零修调；退出使能斜坡归零无突跳。
 *==============================================================================*)

FUNCTION_BLOCK FB_DL_ContourCrossCouple
VAR_INPUT
    fErrX     : LREAL := 0.0;    // X 轴跟随误差 [mm] / X-axis following error [mm]
    fErrY     : LREAL := 0.0;    // Y 轴跟随误差 [mm] / Y-axis following error [mm]
    fDirX     : LREAL := 1.0;    // 轨迹方向向量 X 分量（与 Y 分量构成模 1 向量） [无量纲] / Path direction X component
    fDirY     : LREAL := 0.0;    // 轨迹方向向量 Y 分量 [无量纲] / Path direction Y component
    fKc       : LREAL := 0.5;    // 交叉耦合增益，域 [0,1] [无量纲] / Cross-coupling gain
    fTrimMaxMm: LREAL := 0.5;    // 修调限幅（对称 ±），域 > 0 [mm] / Trim limit [mm]
    fRampMmS  : LREAL := 10.0;   // 修调变化率限，域 > 0 [mm/s] / Trim rate limit [mm/s]
    fCycle    : LREAL := 0.0;    // 扫描周期（<=0 用缺省） [s] / Scan cycle, default used when <= 0
    bEnable   : BOOL := FALSE;   // 使能（FALSE=修调斜坡归零） [-] / Enable, FALSE ramps trim to zero
    bReset    : BOOL := FALSE;   // 复位，上升沿清组态故障锁存 [-] / Reset, rising edge clears config latch
END_VAR
VAR_OUTPUT
    fTrimX  : LREAL;             // X 轴修调注入（已限幅/斜坡） [mm] / X-axis trim injection [mm]
    fTrimY  : LREAL;             // Y 轴修调注入 [mm] / Y-axis trim injection [mm]
    bNoDir  : BOOL;              // 方向向量退化（模过小，零修调直通） [-] / Degenerate direction flag
    bError  : BOOL;              // 组态故障标志（锁存） [-] / Configuration fault flag, latched
END_VAR
VAR
    _fTrimX   : LREAL := 0.0;    // X 修调锁存镜像（斜坡收敛源） / X trim latch mirror
    _fTrimY   : LREAL := 0.0;    // Y 修调锁存镜像 / Y trim latch mirror
    _fTarX    : LREAL;           // 当拍 X 修调目标（斜坡前） [mm] / X trim target before ramp
    _fTarY    : LREAL;           // 当拍 Y 修调目标 [mm] / Y trim target before ramp
    _fEc      : LREAL;           // 当拍轮廓误差 [mm] / Contour error this scan
    _fDen     : LREAL;           // 方向向量模 [无量纲] / Direction vector magnitude
    _fCy      : LREAL;           // 当拍有效周期 [s] / Effective cycle this scan
    _fStep    : LREAL;           // 当拍最大斜坡步长 [mm] / Max ramp step this scan
    _bErrLatch: BOOL;            // 组态故障锁存位（解除沿 = bReset 上升沿） / Latched config fault
    rtReset   : R_TRIG;          // 复位沿实例，段 0 无条件调用 / Reset edge instance
    _bNonFin  : BOOL;            // 输入非有限当拍量 [-] / Non-finite input this scan
    _bNoDir   : BOOL;            // 方向退化当拍量（统一出口映射） / Degenerate direction internal
END_VAR
VAR CONSTANT
    DL_CCC_DIRMIN : LREAL := 1.0E-6;  // 方向向量模下限（防零） [无量纲] / Direction magnitude floor
    DL_CCC_EPS    : LREAL := 0.0;     // 非有限差值判零基准 [-] / Non-finite difference zero base
    DL_CCC_ONE    : LREAL := 1.0;     // 单位常量（增益域上界） [无量纲] / Unit constant
    DL_CCC_CYDEF  : LREAL := 0.01;    // 缺省扫描周期 [s] / Default scan cycle
    DL_CCC_TWO    : LREAL := 2.0;     // 平方指数 [-] / Square exponent base
END_VAR

(* —— 段 0：非有限判 + 组态闸 + 周期派生 + 沿刷新 —— *)
_bNonFin := (fErrX <> fErrX) OR ((fErrX - fErrX) <> DL_CCC_EPS)
         OR (fErrY <> fErrY) OR ((fErrY - fErrY) <> DL_CCC_EPS)
         OR (fDirX <> fDirX) OR ((fDirX - fDirX) <> DL_CCC_EPS)   // 方向 X 非有限（NaN 自反 + Inf 差自减，R79 双判口径对齐，v1.0.1） / Non-finite dir X, dual test
         OR (fDirY <> fDirY) OR ((fDirY - fDirY) <> DL_CCC_EPS);  // 方向 Y 非有限（同双判口径） / Non-finite dir Y, dual test
IF (fKc < 0.0) OR (fKc > DL_CCC_ONE) OR (fTrimMaxMm <= 0.0) OR (fRampMmS <= 0.0) THEN
    _bErrLatch := TRUE;                                     // 组态域闸：锁存（R188 解除沿 = bReset 上升沿） / Config gate: latch
END_IF
IF fCycle > 0.0 THEN
    _fCy := fCycle;                                         // 组态周期有效 / Configured cycle valid
ELSE
    _fCy := DL_CCC_CYDEF;                                   // 周期缺省兜底 / Default cycle fallback
END_IF
_fStep := fRampMmS * _fCy;                                  // 最大斜坡步长 [mm] / Max ramp step
rtReset(CLK := bReset);                                     // 复位沿，每拍必调 / Reset edge, every scan

(* —— 段 1：复位沿 —— *)
IF rtReset.Q THEN
    _bErrLatch := FALSE;                                    // 清组态故障锁存 / Clear config latch
END_IF

(* —— 段 2：轮廓误差与修调目标（故障/退化/非有限分支先行） —— *)
IF _bErrLatch THEN
    _fTarX := 0.0;                                          // 故障安全侧目标零 / Fault safe target zero
    _fTarY := 0.0;                                          // 故障安全侧目标零 / Fault safe target zero
    _bNoDir := FALSE;                                       // 故障期退化标志复位 / Degenerate flag reset
ELSIF _bNonFin THEN
    _fTarX := _fTrimX;                                      // 非有限冻结：目标 = 当前值（保持逼近） / Freeze target to current
    _fTarY := _fTrimY;                                      // 冻结 Y 目标 / Freeze Y target
    _bNoDir := FALSE;                                       // 非有限期不判退化 / No direction judgment
ELSE
    _fDen := SQRT(fDirX * fDirX + fDirY * fDirY);           // 方向向量模（判模后再用，无除零） / Direction magnitude
    IF _fDen < DL_CCC_DIRMIN THEN
        _fTarX := 0.0;                                      // 方向退化：零修调直通（R28 防零） / Degenerate: zero trim
        _fTarY := 0.0;                                      // 零修调 / Zero trim
        _bNoDir := TRUE;                                    // 置退化标志 / Raise degenerate flag
    ELSE
        _fEc := (fErrX * fDirX + fErrY * fDirY) / _fDen;    // 轮廓误差投影（分母模已过闸） / Contour error projection
        _fTarY := fKc * _fEc * fDirX;                       // 垂直分量还给 Y 弱轴 / Vertical component to Y
        _fTarX := -fKc * _fEc * fDirY;                      // 垂直分量还给 X 弱轴（反号） / Vertical component to X, negated
        IF _fTarX > fTrimMaxMm THEN
            _fTarX := fTrimMaxMm;                           // 目标上钳 / Clamp target high
        ELSIF _fTarX < -fTrimMaxMm THEN
            _fTarX := -fTrimMaxMm;                          // 目标下钳 / Clamp target low
        END_IF
        IF _fTarY > fTrimMaxMm THEN
            _fTarY := fTrimMaxMm;                           // 目标上钳 / Clamp target high
        ELSIF _fTarY < -fTrimMaxMm THEN
            _fTarY := -fTrimMaxMm;                          // 目标下钳 / Clamp target low
        END_IF
        _bNoDir := FALSE;                                   // 方向有效 / Direction valid
    END_IF
    IF NOT bEnable THEN
        _fTarX := 0.0;                                      // 未使能目标零（斜坡归零语义，头注释④） / Disabled target zero
        _fTarY := 0.0;                                      // 未使能目标零 / Disabled target zero
    END_IF
END_IF

(* —— 段 3：斜坡逼近（限步长收敛，方向突变/退出使能均无突跳） —— *)
IF _fTarX > (_fTrimX + _fStep) THEN
    _fTrimX := _fTrimX + _fStep;                            // X 正向限步收敛 / X ramp up
ELSIF _fTarX < (_fTrimX - _fStep) THEN
    _fTrimX := _fTrimX - _fStep;                            // X 负向限步收敛 / X ramp down
ELSE
    _fTrimX := _fTarX;                                      // X 步内到达 / X settle
END_IF
IF _fTarY > (_fTrimY + _fStep) THEN
    _fTrimY := _fTrimY + _fStep;                            // Y 正向限步收敛 / Y ramp up
ELSIF _fTarY < (_fTrimY - _fStep) THEN
    _fTrimY := _fTrimY - _fStep;                            // Y 负向限步收敛 / Y ramp down
ELSE
    _fTrimY := _fTarY;                                      // Y 步内到达 / Y settle
END_IF

(* —— 段 4：出口单点映射（名实双出口同源，R191） —— *)
fTrimX := _fTrimX;                                          // X 修调出口 / X trim outlet
fTrimY := _fTrimY;                                          // Y 修调出口 / Y trim outlet
bNoDir := _bNoDir AND (NOT _bErrLatch);                     // 退化标志出口（故障期复位） / Degenerate outlet
bError := _bErrLatch;                                       // 故障标志出口 / Error flag outlet

END_FUNCTION_BLOCK

(* ---- FB_DL_CrankKinFwd.st ---- *)
// FB_DL_CrankKinFwd v1.0.0
// 开源溯源：self-cleanroom / 公开运动学公式（曲柄滑块机构）
(*
  道莅工业代码库 | DL_Motion | FB_DL_CrankKinFwd
  版本: 1.0.0 | 日期: 2026-11-23 | 轮次: R75
  功能: 曲柄滑块机构正运动学：曲柄角 θ → 滑块位移 x = r·cosθ +
        sqrt(L² − r²·sin²θ)；附角速度输入时的滑块速度解析导数
        ẋ = −ω·r·sinθ·(1 + r·cosθ/sqrt(L² − r²·sin²θ))
  邻件关系: robot 族（监视/抓取验证）与本件无运动学属主重叠；并联件
            FB_DL_DeltaRobotIk 为逆解（末端→关节），本件为正解
            （关节→末端），方向互补
  机构约束: 连杆长 L 必须大于曲柄半径 r（L−r > 容差），否则机构无法
            整周回转，判组态故障拒算
*)
FUNCTION_BLOCK FB_DL_CrankKinFwd
VAR_INPUT
    bEnable    : BOOL := FALSE;             // 使能（FALSE 输出保持零）/ Enable
    fCrankDeg  : REAL := 0.0;               // 曲柄角 θ [deg]，0=TDC，域 ±1E6 / Crank angle [deg], 0 at TDC
    fOmegaRadS : REAL := 0.0;               // 曲柄角速度 ω [rad/s]，0 时速度输出零 / Crank angular velocity [rad/s]
    fCrankR    : REAL := 25.0;              // 曲柄半径 r [mm]，域 > 0 / Crank radius [mm]
    fRodL      : REAL := 100.0;             // 连杆长 L [mm]，域 > r + 容差 / Connecting rod length [mm]
    fEps       : REAL := 1.0E-6;            // 判零/判界容差 [mm] / Tolerance [mm]
END_VAR
VAR_OUTPUT
    fSliderPos : REAL;                      // 滑块位移（距曲轴心）[mm] / Slider position from crank center [mm]
    fSliderVel : REAL;                      // 滑块速度 [mm/s] / Slider velocity [mm/s]
    bValid     : BOOL;                      // 结果有效回执 [-] / Result validity receipt
    bError     : BOOL;                      // 故障标志（机构约束违反）/ Fault flag (mechanism constraint violated)
    uErrorId   : UDINT;                     // 事件码，0 = 无事件；16#0002_2701 = 组态非法 / Event code
END_VAR
VAR
    fThetaRad  : REAL;                      // 弧度角 [rad] / Angle in radians
    fSinT      : REAL;                      // sin θ [1] / Sine of angle
    fCosT      : REAL;                      // cos θ [1] / Cosine of angle
    fRad2      : REAL;                      // 根号内 L² − r²sin²θ [mm²] / Radicand
    fRoot      : REAL;                      // sqrt 根号值 [mm] / Square root value
    fRr        : REAL;                      // 曲柄半径平方 [mm²] / Radius squared
    fLr        : REAL;                      // 连杆长平方 [mm²] / Rod length squared
END_VAR

// —— 段 0：全路径缺省 —— //
fSliderPos := 0.0;                       // 位移缺省零 / Position default zero
fSliderVel := 0.0;                       // 速度缺省零 / Velocity default zero
bValid := FALSE;                         // 有效回执预清 / Validity preset
bError := FALSE;                         // 故障预清（约束违反路径置位）/ Fault preset
uErrorId := 16#0000;                     // 事件码预清 / Event code preset

// —— 段 1：机构约束闸与输入闸 —— //
IF (fCrankR <> fCrankR) OR (fRodL <> fRodL) OR (fCrankDeg <> fCrankDeg) OR (fOmegaRadS <> fOmegaRadS) THEN
    bError := TRUE;                      // 故障级：输入含 NaN / Fault level: NaN input
    uErrorId := 16#0002_2701;            // 故障码（27xx 步进）/ Fault code
    RETURN;
END_IF
IF (fCrankR <= fEps) OR (fRodL <= fCrankR + fEps) THEN
    bError := TRUE;                      // 故障级：曲柄非正或连杆不长于曲柄（机构约束）/ Fault level: mechanism constraint
    uErrorId := 16#0002_2701;            // 同码段复用（R90 不加码：同属组态非法）/ Same code family
    RETURN;
END_IF
bValid := TRUE;                          // 组态与输入均有效 / Validity receipt

// —— 段 2：使能门控 —— //
IF NOT bEnable THEN
    fSliderPos := 0.0;                   // 失能输出零 / Disabled zero output
    fSliderVel := 0.0;                   // 速度零 / Velocity zero
    RETURN;                              // 失能不计算 / No computation when disabled
END_IF

// —— 段 3：正运动学主计算 —— //
fThetaRad := fCrankDeg * 0.017453292519943295;   // 角度转弧度（π/180 常数）/ Deg to rad
fSinT := SIN(fThetaRad);                 // sin θ / Sine
fCosT := COS(fThetaRad);                 // cos θ / Cosine
fRr := fCrankR * fCrankR;                // r² [mm²] / Radius squared
fLr := fRodL * fRodL;                    // L² [mm²] / Rod length squared
fRad2 := fLr - fRr * fSinT * fSinT;      // L² − r²sin²θ（≥ L² − r² > 0 已过闸）/ Radicand, positive by gate
fRoot := SQRT(fRad2);                    // 根号值 [mm] / Root value
fSliderPos := fCrankR * fCosT + fRoot;   // 滑块位移 x = r·cosθ + sqrt(...) / Slider position
fSliderVel := -fOmegaRadS * fCrankR * fSinT * (1.0 + fCrankR * fCosT / fRoot);   // 解析速度 [mm/s]（fRoot > 0 已过闸）/ Analytic velocity
END_FUNCTION_BLOCK

(* ---- FB_DL_DeltaRobotIk.st ---- *)
(*
  道莅工业代码库 | DL_Motion | FB_DL_DeltaRobotIk
  版本: 1.0.0 | 日期: 2026-11-23 | 轮次: R75
  开源溯源: self-cleanroom（无外部来源；Delta 并联机构闭式逆解为公开几何推导，
            本件由解析几何独立推导实现，零代码行复制）
  功能: 三臂并联三角洲机器人逆运动学——末端 XYZ [mm] → 三臂上臂关节角 [°]
        （相对水平面，肘下主解分支），含行程奇异性闸与可达性闸。
  兼容性: CODESYS 3.5 / TwinCAT 3 / 汇川 InoProShop；仅依赖标准 SQRT/ABS/ACOS/ATAN，零厂商私有库
  接口: 输入末端 XYZ 与机构四参数（基座半径/动平台半径/上臂长/前臂长）+ 上臂角限位；
        输出三臂角 fTheta1Deg~fTheta3Deg [°]、bReachOk、eErr。变换型 FB（无相位机，
        每拍独立全量重算，无跨周期状态），无 TON/R_TRIG 实例。
  码表: 16#0004_0369 故障级：参数非法（半径/臂长/限位角非法或末端坐标非有限）
        16#0004_036A 故障级：目标不可达（侧偏超限无解/三角函数域越界/上臂角超行程）
        码段说明：0004 段故障子带 03xx，槽位经全库实扫空闲。
  边界: ① 逆解方程：uXr*cosφ - fZ*sinφ = C（C = -(K²-Lu²-X²-z²)/(2Lu)），
        化为 R·cos(φ+α) 求解，α 由 ATAN 加象限修正手构（不用方言 ATAN2）；
        ② 侧向偏移使 K² = Lf²-b² < 0 判不可达（奇异性闸前置）；
        ③ 所有除法分母先闸（2Lu 由参数闸 >0 证明，R 由 EPS 下限闸，uXr 由 ABS<EPS 闸）；
        ④ 上臂角限位 |φ| > fPhiMaxDeg 判行程越界；
        ⑤ 任一臂不可达 → 三臂输出全零（不输出部分解）；⑥ 零全局耦合。
  邻件比对: robot 族仅监视/抓取验证件在册，无运动学逆解属主（R75 §3 留痕）。
  修订历史: 2026-11-23 v1.0.0 R75 首版（复杂件批 B1 · C03）
*)

FUNCTION_BLOCK FB_DL_DeltaRobotIk
VAR_INPUT
    fX         : LREAL := 0.0;    // 末端 X 坐标 [mm] | End-effector X coordinate
    fY         : LREAL := 0.0;    // 末端 Y 坐标 [mm] | End-effector Y coordinate
    fZ         : LREAL := 0.0;    // 末端 Z 坐标（基座平面上方为正）[mm] | End-effector Z coordinate, positive above base plane
    fRBase     : LREAL := 200.0;  // 基座等边三角形半径（肩关节分布圆），域 > 0 [mm] | Base triangle radius
    fRPlat     : LREAL := 50.0;   // 动平台等边三角形半径（腕关节分布圆），域 > 0 [mm] | Platform triangle radius
    fArmLen    : LREAL := 100.0;  // 上臂长度，域 > 0 [mm] | Upper arm length
    fForeLen   : LREAL := 250.0;  // 前臂（从动杆）长度，域 > 0 [mm] | Forearm length
    fPhiMaxDeg : LREAL := 80.0;   // 上臂角限位幅值，域 (0, 180) [°] | Upper arm angle travel limit
END_VAR
VAR_OUTPUT
    fTheta1Deg : LREAL;           // 臂 1 上臂关节角（方位 0°，相对水平面）[°] | Arm 1 upper joint angle at azimuth 0 deg
    fTheta2Deg : LREAL;           // 臂 2 上臂关节角（方位 120°）[°] | Arm 2 upper joint angle at azimuth 120 deg
    fTheta3Deg : LREAL;           // 臂 3 上臂关节角（方位 240°）[°] | Arm 3 upper joint angle at azimuth 240 deg
    bReachOk   : BOOL;            // 可达且行程内 [-] | Reachable and within travel
    eErr       : UDINT;           // 错误码，0 = 无错 | Error code, 0 = none
END_VAR
VAR
    aTheta   : ARRAY[1..3] OF LREAL;  // 三臂角暂存（出口统一映射）[°] | Per-arm angle staging
    uPsiCos  : LREAL;                 // 当前臂方位角余弦 [-] | Current arm azimuth cosine
    uPsiSin  : LREAL;                 // 当前臂方位角正弦 [-] | Current arm azimuth sine
    uXr      : LREAL;                 // 目标在臂平面内的径向差 [mm] | Radial offset in arm plane
    uLat     : LREAL;                 // 目标侧向偏移（离臂平面）[mm] | Lateral offset out of arm plane
    uK2      : LREAL;                 // 可达半径平方 K² [mm²] | Squared reachable radius
    uK       : LREAL;                 // 可达半径 K [mm] | Reachable radius
    uM       : LREAL;                 // 化简常数 M [mm] | Reduced constant
    uR       : LREAL;                 // 径向-高度合成半径 R [mm] | Combined radial-height radius
    uCosv    : LREAL;                 // cos(φ+α) 候补 [-] | cos of phi plus alpha candidate
    uAlpha   : LREAL;                 // 象限修正后的 α [rad] | Quadrant-corrected alpha
    uPhi     : LREAL;                 // 上臂角主解 [rad] | Upper arm angle primary solution
    i        : INT;                   // 臂序号游标 | Arm index cursor
    bOk      : BOOL;                  // 全程可达标志 [-] | All arms reachable flag
END_VAR
VAR CONSTANT
    DL_DRI_PI     : LREAL := 3.14159265358979;    // 圆周率 | Pi
    DL_DRI_EPS    : LREAL := 1.0E-9;              // 退化判定容差 [mm] | Degeneracy tolerance
    DL_DRI_RAD2DEG: LREAL := 57.29577951308232;   // 弧度转角度因子 | Rad to deg factor
    DL_DRI_ERR_PAR: UDINT := 16#0004_0369;        // 参数非法码 | Illegal parameter code
    DL_DRI_ERR_REA: UDINT := 16#0004_036A;        // 不可达码 | Unreachable code
END_VAR

(* —— 段 0：输出缺省全赋值（全路径覆盖） —— *)
aTheta[1] := 0.0;                       // 臂 1 暂存清零（防御） / Arm 1 staging cleared
aTheta[2] := 0.0;                       // 臂 2 暂存清零（防御） / Arm 2 staging cleared
aTheta[3] := 0.0;                       // 臂 3 暂存清零（防御） / Arm 3 staging cleared
bReachOk := FALSE;                      // 可达标志预置 FALSE / Reach flag preset FALSE
eErr := 0;                              // 错误码缺省 / Error default

(* —— 段 1：输入与机构参数域闸 —— *)
bOk := TRUE;                            // 可达标志初值 / Reach flag init
IF (fX <> fX) OR (fY <> fY) OR (fZ <> fZ)
   OR (fRBase <> fRBase) OR (fRPlat <> fRPlat) OR (fArmLen <> fArmLen)
   OR (fForeLen <> fForeLen) OR (fPhiMaxDeg <> fPhiMaxDeg) THEN
    bOk := FALSE;                       // 任一输入非有限 / Any non-finite input
    eErr := DL_DRI_ERR_PAR;             // 参数非法码 / Parameter code
END_IF
IF bOk AND ((fRBase <= 0.0) OR (fRPlat <= 0.0) OR (fArmLen <= 0.0)
         OR (fForeLen <= 0.0) OR (fPhiMaxDeg <= 0.0) OR (fPhiMaxDeg >= 180.0)) THEN
    bOk := FALSE;                       // 机构参数越域 / Mechanism parameters out of domain
    eErr := DL_DRI_ERR_PAR;             // 参数非法码 / Parameter code
END_IF

(* —— 段 2：三臂逆解主循环（肘下主解分支；任一臂失败即全件失败） —— *)
IF bOk THEN
    FOR i := 1 TO 3 DO
        // 方位角常量展开（免数组字面量初始化，跨平台安全）/ Azimuth constants unrolled
        CASE i OF
        1:  uPsiCos := 1.0;                                             // 臂 1 方位 0° | Arm 1 azimuth 0 deg
            uPsiSin := 0.0;
        2:  uPsiCos := -0.5;                                            // 臂 2 方位 120° | Arm 2 azimuth 120 deg
            uPsiSin := 0.866025403784439;
        3:  uPsiCos := -0.5;                                            // 臂 3 方位 240° | Arm 3 azimuth 240 deg
            uPsiSin := -0.866025403784439;
        ELSE
            uPsiCos := 1.0;                                             // 不可达分支兜底（循环上界已闸 1..3） | Unreachable fallback
            uPsiSin := 0.0;
        END_CASE

        // 几何量：径向差 / 侧偏 / 可达半径平方
        uXr := fX * uPsiCos + fY * uPsiSin - (fRBase - fRPlat);         // 径向差 X = x·cosψ + y·sinψ - (Rb-Rp) / Radial offset
        uLat := -fX * uPsiSin + fY * uPsiCos;                           // 侧偏 b = -x·sinψ + y·cosψ / Lateral offset
        uK2 := fForeLen * fForeLen - uLat * uLat;                       // K² = Lf² - b² / Squared reachable radius
        IF uK2 < 0.0 THEN
            bOk := FALSE;                                               // 侧偏超限无解（奇异性闸） / Lateral offset beyond reach
            eErr := DL_DRI_ERR_REA;                                     // 不可达码 / Unreachable code
        ELSE
            uK := SQRT(uK2);                                            // 可达半径 K ≥ 0 / Reachable radius
            uM := (uK2 - fArmLen * fArmLen - uXr * uXr - fZ * fZ)
               / (2.0 * fArmLen);                                       // M = (K²-Lu²-X²-z²)/(2Lu)，分母由参数闸 >0 / Reduced constant, denominator proven
            uR := SQRT(uXr * uXr + fZ * fZ);                            // 合成半径 R = √(X²+z²) / Combined radius
            IF uR < DL_DRI_EPS THEN
                IF ABS(uM) < DL_DRI_EPS THEN
                    uPhi := 0.0;                                        // 退化同心且 M≈0：φ=0 / Degenerate concentric, phi = 0
                ELSE
                    bOk := FALSE;                                       // 退化且无解 / Degenerate unsolvable
                    eErr := DL_DRI_ERR_REA;
                END_IF
            ELSE
                uCosv := -uM / uR;                                      // cos(φ+α) = -M/R，分母已闸 R > EPS / Cosine candidate, denominator gated
                IF ABS(uCosv) > 1.0 THEN
                    bOk := FALSE;                                       // 反余弦定义域越界 = 不可达 / acos domain violated, unreachable
                    eErr := DL_DRI_ERR_REA;
                ELSE
                    // α = atan2(fZ, uXr) 手构象限修正（不用方言 ATAN2）/ Manual atan2 with quadrant fix
                    IF ABS(uXr) < DL_DRI_EPS THEN
                        IF fZ >= 0.0 THEN
                            uAlpha := 0.5 * DL_DRI_PI;                  // X≈0 且 z≥0：α=+π/2 | X near zero, z non-negative
                        ELSE
                            uAlpha := -0.5 * DL_DRI_PI;                 // X≈0 且 z<0：α=-π/2 | X near zero, z negative
                        END_IF
                    ELSE
                        uAlpha := ATAN(fZ / uXr);                       // 分母 ABS(uXr) >= EPS 已闸 / Denominator gated
                        IF uXr < 0.0 THEN
                            IF fZ >= 0.0 THEN
                                uAlpha := uAlpha + DL_DRI_PI;           // 第二象限修正 | Second quadrant fix
                            ELSE
                                uAlpha := uAlpha - DL_DRI_PI;           // 第三象限修正 | Third quadrant fix
                            END_IF
                        END_IF
                    END_IF
                    uPhi := ACOS(uCosv) - uAlpha;                       // 肘下主解：φ = acos(-M/R) - α / Elbow-down primary branch
                END_IF
            END_IF
        END_IF

        IF bOk THEN
            IF ABS(uPhi * DL_DRI_RAD2DEG) > fPhiMaxDeg THEN
                bOk := FALSE;                                           // 上臂角超行程限位 / Upper arm angle beyond travel
                eErr := DL_DRI_ERR_REA;                                 // 不可达码（行程越界归并） / Unreachable code folded
            ELSE
                aTheta[i] := uPhi * DL_DRI_RAD2DEG;                     // 弧度转角度入暂存 / Rad to deg into staging
            END_IF
        END_IF
    END_FOR
END_IF

(* —— 段 3：出口单点映射（失败全零输出，不输出部分解） —— *)
fTheta1Deg := aTheta[1];                // 臂 1 角出口 [°] / Arm 1 angle outlet
fTheta2Deg := aTheta[2];                // 臂 2 角出口 [°] / Arm 2 angle outlet
fTheta3Deg := aTheta[3];                // 臂 3 角出口 [°] / Arm 3 angle outlet
bReachOk := bOk;                        // 可达出口（名实同源） / Reach outlet

END_FUNCTION_BLOCK
